        IF NOT stCmd.bEnable THEN
            // Route disable through STOPPING so MC_Stop runs first. If torque was
            // applied the axis is still in CST (torque) mode after Stop Torque;
            // MC_Stop performs the CST->position changeover and decelerates to a
            // real standstill BEFORE MC_Power drops. Withdrawing controller enable
            // straight from CST tripped NC 0x4260 (enable removed while the axis
            // was still positioning). STOPPING -> fbStop.Done -> DISABLED (SEL on
            // bEnable). Brief position hold during the decel, then power-off leaves
            // the motor free. (MOVING already disables via STOPPING; this makes
            // READY consistent. A normal idle disable just no-op-stops through it.)
            eState := E_MotorState.STOPPING;
        ELSIF fbPower.Error THEN
            eState := E_MotorState.ERROR;
        ELSIF rtStop.Q THEN
            eState := E_MotorState.STOPPING;
        ELSIF rtHome.Q THEN
            eState := E_MotorState.HOMING;
        ELSIF rtExecuteMove.Q THEN
            bMoveLatch := TRUE;
            eState     := E_MotorState.MOVING;
        END_IF

    E_MotorState.MOVING:
        IF NOT stCmd.bEnable OR rtStop.Q THEN
            bMoveLatch := FALSE;
            eState     := E_MotorState.STOPPING;

        ELSIF stCmd.eControlMode = E_ControlMode.POSITION THEN
            IF stCmd.bRelative THEN
                IF fbMoveRel.Busy  THEN bMoveLatch := FALSE; END_IF
                IF fbMoveRel.Done  THEN eState := E_MotorState.READY; END_IF
                IF fbMoveRel.Error THEN eState := E_MotorState.ERROR; END_IF
            ELSE
                IF fbMoveAbs.Busy  THEN bMoveLatch := FALSE; END_IF
                IF fbMoveAbs.Done  THEN eState := E_MotorState.READY; END_IF
                IF fbMoveAbs.Error THEN eState := E_MotorState.ERROR; END_IF
            END_IF

        ELSIF stCmd.eControlMode = E_ControlMode.VELOCITY THEN
            IF stCmd.fTargetVelocity <> fPrevVelocity THEN
                fPrevVelocity := stCmd.fTargetVelocity;
                bMoveLatch    := TRUE;
            END_IF
            IF fbMoveVel.Busy  THEN bMoveLatch := FALSE; END_IF
            IF fbMoveVel.Error THEN eState := E_MotorState.ERROR; END_IF

        ELSE
            eState := E_MotorState.READY;
        END_IF

    E_MotorState.STOPPING:
        IF fbStop.Error THEN
            eState := E_MotorState.ERROR;
        ELSIF fbStop.Done THEN
            eState := SEL(stCmd.bEnable, E_MotorState.DISABLED, E_MotorState.READY);
        END_IF

    E_MotorState.HOMING:
        fbHome(Axis := Axis, Execute := TRUE, HomingMode := MC_DefaultHoming);
        IF fbHome.Error THEN
            eState := E_MotorState.ERROR;
        ELSIF fbHome.Done THEN
            stStatus.bHomingDone := TRUE;
            eState               := E_MotorState.READY;
        END_IF

    E_MotorState.ERROR:
        IF rtResetError.Q THEN
            // Sequenced recovery: clear the DRIVE fault first (SoE S-0-0099),
            // give the drive a settle gap, THEN reset the NC axis against the
            // healthy drive. Sequenced on COMPLETION (Busy/Done), not timers.
            bSoeResetExec := TRUE;
            nResetStage   := 1;
            eState        := E_MotorState.RESETTING;
        END_IF

    E_MotorState.RESETTING:
        // Whole-sequence watchdog: if any stage hangs (e.g. a latch that never
        // clears), give up and go BACK TO ERROR — visible failure, another
        // reset press retries. Without this a stuck stage is unrecoverable
        // until a PLC restart.
        tonResetGuard(IN := TRUE, PT := T_RESET_GUARD);
        IF tonResetGuard.Q THEN
            tonResetGuard(IN := FALSE);
            bSoeResetExec := FALSE;
            bNcResetExec  := FALSE;
            nResetStage   := 0;
            eState        := E_MotorState.ERROR;
        END_IF
        CASE nResetStage OF
            1:  // SoE drive reset running — the latch self-clears when the
                // FB's Busy falls (done) or it errors/times out (10 s)
                IF NOT bSoeResetExec THEN
                    tonSettle(IN := FALSE);
                    nResetStage := 2;
                END_IF
            2:  // settle: let the drive's state machine come back up before
                // the NC touches it
                tonSettle(IN := TRUE, PT := T_RESET_SETTLE);
                IF tonSettle.Q THEN
                    tonSettle(IN := FALSE);
                    bNcResetExec := TRUE;
                    nResetStage  := 3;
                END_IF
            3:  // NC axis reset — latch self-clears on Done/Error
                IF NOT bNcResetExec THEN
                    tonResetGuard(IN := FALSE);
                    stStatus.bError   := FALSE;
                    stStatus.nErrorID := 0;
                    nResetStage       := 0;
                    eState            := E_MotorState.DISABLED;
                END_IF
        END_CASE

END_CASE

//----------------------------------------------------------------------
// STATUS OUTPUTS
//----------------------------------------------------------------------
stStatus.eState       := eState;
stStatus.eControlMode := stCmd.eControlMode;
stStatus.nResetStage  := nResetStage;
stStatus.bEnabled     := fbPower.Status;
stStatus.bMoving      := fbMoveAbs.Busy OR fbMoveRel.Busy OR fbMoveVel.Busy;
stStatus.bAtTarget    := fbMoveAbs.Done OR fbMoveRel.Done OR fbMoveVel.InVelocity;
// Error status sourced from the NC axis ErrorCode — the authoritative, PERSISTENT
// fault: set on any axis fault and HELD until MC_Reset. The MC-block .Error outputs
// are transient (they clear the moment a block's Execute drops or the axis
// disables), so the old MC-block-only bError usually went FALSE before the app
// polled and the error never reached the GUI (nErrorID lingered with bError=FALSE).
// Keep the block errors OR'd in; fall back to their ErrorID only when the axis has
// no code of its own; clear when truly error-free so a stale code can't linger.
stStatus.bError := (Axis.NcToPlc.ErrorCode <> 0)
                OR fbPower.Error   OR fbMoveAbs.Error OR fbMoveRel.Error
                OR fbMoveVel.Error OR fbStop.Error    OR fbHome.Error;

IF Axis.NcToPlc.ErrorCode <> 0 THEN
    stStatus.nErrorID := Axis.NcToPlc.ErrorCode;
ELSIF stStatus.bError THEN
    stStatus.nErrorID := SEL(fbPower.Error,   0, fbPower.ErrorID)
                       + SEL(fbMoveAbs.Error, 0, fbMoveAbs.ErrorID)
                       + SEL(fbMoveRel.Error, 0, fbMoveRel.ErrorID)
                       + SEL(fbMoveVel.Error, 0, fbMoveVel.ErrorID)
                       + SEL(fbStop.Error,    0, fbStop.ErrorID)
                       + SEL(fbHome.Error,    0, fbHome.ErrorID);
ELSE
    stStatus.nErrorID := 0;
END_IF

stStatus.fActPosition := Axis.NcToPlc.ActPos;
stStatus.fActVelocity := Axis.NcToPlc.ActVelo;
stStatus.fActTorque   := INT_TO_LREAL(nActTorque_Raw) / 10.0;
stStatus.nTimestamp   := ULINT_TO_UDINT(F_GetSystemTime() / 10000);

END_FUNCTION_BLOCK

// ---- POUs/FB_TorqueControl.TcPOU
FUNCTION_BLOCK FB_TorqueControl
VAR_IN_OUT
    Axis            : AXIS_REF;         // Must be VAR_IN_OUT — passed by reference
END_VAR

VAR_INPUT
    stCmd           : ST_MotorCommand;  // Read from GVL_Commands
    bAxisReady      : BOOL;             // gate: only stream torque while the axis is READY
END_VAR

VAR_OUTPUT
    stStatus        : ST_MotorStatus;   // Written to GVL_Status
END_VAR

VAR
    fbTorqueCtrl    : MC_TorqueControl;
    rtExecute       : R_TRIG;
END_VAR

// Rising edge on bTorqueExecute triggers MC_TorqueControl
rtExecute(CLK := stCmd.bTorqueExecute);

// Gate Execute on READY: torque must never be commanded on a DISABLED/ERROR/
// RESETTING axis. This also drops Execute on a fault (READY->ERROR), which
// clears MC_TorqueControl's latched Error, and prevents the reset "bounce"
// where torque errors on the just-disabled axis and re-stamps the fault.
fbTorqueCtrl(
    Axis              := Axis,
    Execute           := stCmd.bTorqueExecute AND bAxisReady,
    ContinuousUpdate  := TRUE,
    Relative          := FALSE,
    Torque            := stCmd.fTargetTorque,
    TorqueRamp        := stCmd.fTorqueRamp,
    VelocityLimitHigh := stCmd.fTorqueVelLimitHigh,
    VelocityLimitLow  := stCmd.fTorqueVelLimitLow,
    BufferMode        := MC_Aborting
);

// Write ONLY torque fields back — do not overwrite position/velocity status
stStatus.bTorqueActive   := fbTorqueCtrl.Active;
stStatus.bTorqueInTorque := fbTorqueCtrl.InTorque;

// Reflect the LIVE torque-FB error. This was set-only (no ELSE), so once a
// torque fault set bError it stayed latched forever and PRG_Motion's set-only
// copy re-stamped it onto the status mirror every scan — the motor recovered
// but bError/nErrorID never cleared. With Execute gated off on !READY, a reset
// clears MC_TorqueControl.Error and this ELSE then clears the mirror. A REAL,
// persistent torque fault keeps fbTorqueCtrl.Error TRUE, so it is not masked.
IF fbTorqueCtrl.Error THEN
    stStatus.bError   := TRUE;
    stStatus.nErrorID := fbTorqueCtrl.ErrorId;
ELSE
    stStatus.bError   := FALSE;
    stStatus.nErrorID := 0;
END_IF

END_FUNCTION_BLOCK

// ---- POUs/FB_IOHandler.TcPOU
FUNCTION_BLOCK FB_IOHandler
VAR_INPUT
    // Raw digital input byte — link this to your EL1008 terminal in XAE
    nRawDigitalIn   : BYTE;

    // Raw analog input values — link to EL3002 channels in XAE
    nRawAnalogIn_Ch1 : INT;
    nRawAnalogIn_Ch2 : INT;

    // Analog scaling — set once from MAIN or leave as defaults
    fAnalogIn_Scale_Ch1  : LREAL := 10.0;   // full-scale [V or mA]
    fAnalogIn_Scale_Ch2  : LREAL := 10.0;
    fAnalogOut_Scale_Ch1 : LREAL := 10.0;
    fAnalogOut_Scale_Ch2 : LREAL := 10.0;
END_VAR

VAR_OUTPUT
    // Packed digital output byte — link this to your EL2008 terminal in XAE
    nRawDigitalOut  : BYTE;

    // Raw analog output values — link to EL4002 channels in XAE
    nRawAnalogOut_Ch1 : INT;
    nRawAnalogOut_Ch2 : INT;
END_VAR

VAR_IN_OUT
    // Shared IO struct — same instance passed in from MAIN and GVL_IO
    stIO : ST_IOData;
END_VAR

//======================================================================
// DIGITAL INPUTS — unpack raw byte into named booleans
//======================================================================
stIO.bDI_EmergencyStop  := nRawDigitalIn.0;
stIO.bDI_HomeSensor_M1  := nRawDigitalIn.1;
stIO.bDI_HomeSensor_M2  := nRawDigitalIn.2;
stIO.bDI_LimitPos_M1    := nRawDigitalIn.3;
stIO.bDI_LimitNeg_M1    := nRawDigitalIn.4;
stIO.bDI_LimitPos_M2    := nRawDigitalIn.5;
stIO.bDI_LimitNeg_M2    := nRawDigitalIn.6;
stIO.bDI_UserInput1     := nRawDigitalIn.7;

// Mirror raw byte for Python diagnostics
stIO.nDigitalInputs     := nRawDigitalIn;

//======================================================================
// ANALOG INPUTS — scale INT [-32768..32767] → engineering units
// Formula: value = (raw / 32767.0) * full_scale
//======================================================================
stIO.fAnalogIn_Ch1      := (INT_TO_LREAL(nRawAnalogIn_Ch1) / 32767.0)
                            * fAnalogIn_Scale_Ch1;
stIO.fAnalogIn_Ch2      := (INT_TO_LREAL(nRawAnalogIn_Ch2) / 32767.0)
                            * fAnalogIn_Scale_Ch2;
stIO.nAnalogIn_Raw_Ch1  := nRawAnalogIn_Ch1;
stIO.nAnalogIn_Raw_Ch2  := nRawAnalogIn_Ch2;

//======================================================================
// DIGITAL OUTPUTS — pack named booleans into raw byte for EL2008
//======================================================================
nRawDigitalOut.0 := stIO.bDO_BrakeRelease_M1;
nRawDigitalOut.1 := stIO.bDO_BrakeRelease_M2;
nRawDigitalOut.2 := stIO.bDO_StatusLED_Green;
nRawDigitalOut.3 := stIO.bDO_StatusLED_Red;
nRawDigitalOut.4 := stIO.bDO_UserOutput1;
nRawDigitalOut.5 := stIO.bDO_UserOutput2;

// Mirror packed byte back into struct for Python readback
stIO.nDigitalOutputs    := nRawDigitalOut;

//======================================================================
// ANALOG OUTPUTS — scale engineering units → INT [-32767..32767]
// Formula: raw = CLAMP(value / full_scale, -1.0, 1.0) * 32767
// Python writes fAnalogOut_Ch1/2 into GVL_IO.stIO, FB reads them here
//======================================================================
stIO.nAnalogOut_Raw_Ch1 := LREAL_TO_INT(
    LIMIT(-32767.0,
          (stIO.fAnalogOut_Ch1 / fAnalogOut_Scale_Ch1) * 32767.0,
          32767.0));

stIO.nAnalogOut_Raw_Ch2 := LREAL_TO_INT(
    LIMIT(-32767.0,
          (stIO.fAnalogOut_Ch2 / fAnalogOut_Scale_Ch2) * 32767.0,
          32767.0));

nRawAnalogOut_Ch1 := stIO.nAnalogOut_Raw_Ch1;
nRawAnalogOut_Ch2 := stIO.nAnalogOut_Raw_Ch2;

END_FUNCTION_BLOCK

// ---- POUs/FB_EncoderHandler.TcPOU
FUNCTION_BLOCK FB_EncoderHandler
VAR_IN_OUT
    stEncoder           : ST_EncoderData;
END_VAR

VAR_INPUT
    fCountsPerUnit      : LREAL := 1.0;
END_VAR

VAR
    nStatusWord_Raw      AT %I* : WORD;
    nCounterValue_Raw    AT %I* : DWORD;
    nFrequencyValue_Raw  AT %I* : DWORD;
    nState_Raw           AT %I* : BYTE;

    nSetCounterValue_Raw AT %Q* : DWORD;
    nControlWord_Raw     AT %Q* : WORD;

    rtSetCounter        : R_TRIG;
    rtZeroPosition      : R_TRIG;
END_VAR

//----------------------------------------------------------------------
// READ INPUTS
//----------------------------------------------------------------------
stEncoder.nStatusWord     := nStatusWord_Raw;
stEncoder.nCounterValue   := nCounterValue_Raw;
stEncoder.nFrequencyValue := nFrequencyValue_Raw;
stEncoder.nState          := nState_Raw;

stEncoder.bInputA           := nStatusWord_Raw.0;
stEncoder.bInputB           := nStatusWord_Raw.1;
stEncoder.bInputC           := nStatusWord_Raw.2;
stEncoder.bCounterUnderflow := nStatusWord_Raw.4;
stEncoder.bCounterOverflow  := nStatusWord_Raw.5;
stEncoder.bLatchValid       := nStatusWord_Raw.8;
stEncoder.bError            := nStatusWord_Raw.14;

IF fCountsPerUnit <> 0 THEN
    stEncoder.fPosition := DWORD_TO_LREAL(nCounterValue_Raw) / fCountsPerUnit;
END_IF

//----------------------------------------------------------------------
// WRITE OUTPUTS
//----------------------------------------------------------------------
rtSetCounter  (CLK := stEncoder.bSetCounter);
rtZeroPosition(CLK := stEncoder.bZeroPosition);

IF rtZeroPosition.Q THEN
    stEncoder.nSetCounterValue := 0;
    nSetCounterValue_Raw       := 0;
    nControlWord_Raw.2         := TRUE;   // bit 2 = 0x7000:03 Set counter
ELSIF rtSetCounter.Q THEN
    nSetCounterValue_Raw       := stEncoder.nSetCounterValue;
    nControlWord_Raw.2         := TRUE;
ELSE
    nControlWord_Raw.2         := FALSE;
END_IF

END_FUNCTION_BLOCK

// ---- POUs/FB_AnalogInHandler.TcPOU
FUNCTION_BLOCK FB_AnalogInHandler
VAR_IN_OUT
    stAnalogIn      : ST_AnalogInData;  // Shared with GVL_AnalogIn
END_VAR

VAR
    //--- EL3702 PDO inputs — oversampling x5 per channel ---
    // Each sample is a signed INT [-32768 to 32767]
    // AT %I* — linked in XAE instance tree to EL3702 PDO channels
    nCh1_S1     AT %I* : INT;   // Ch1 sample 1
    nCh1_S2     AT %I* : INT;   // Ch1 sample 2
    nCh1_S3     AT %I* : INT;   // Ch1 sample 3
    nCh1_S4     AT %I* : INT;   // Ch1 sample 4
    nCh1_S5     AT %I* : INT;   // Ch1 sample 5

    nCh2_S1     AT %I* : INT;   // Ch2 sample 1
    nCh2_S2     AT %I* : INT;   // Ch2 sample 2
    nCh2_S3     AT %I* : INT;   // Ch2 sample 3
    nCh2_S4     AT %I* : INT;   // Ch2 sample 4
    nCh2_S5     AT %I* : INT;   // Ch2 sample 5

    //--- Internal ---
    fCh1_Sum    : LREAL;
    fCh2_Sum    : LREAL;
    fScale      : LREAL;
END_VAR

//----------------------------------------------------------------------
// STORE RAW SAMPLES INTO STRUCT
//----------------------------------------------------------------------
stAnalogIn.nCh1_Sample[1] := nCh1_S1;
stAnalogIn.nCh1_Sample[2] := nCh1_S2;
stAnalogIn.nCh1_Sample[3] := nCh1_S3;
stAnalogIn.nCh1_Sample[4] := nCh1_S4;
stAnalogIn.nCh1_Sample[5] := nCh1_S5;

stAnalogIn.nCh2_Sample[1] := nCh2_S1;
stAnalogIn.nCh2_Sample[2] := nCh2_S2;
stAnalogIn.nCh2_Sample[3] := nCh2_S3;
stAnalogIn.nCh2_Sample[4] := nCh2_S4;
stAnalogIn.nCh2_Sample[5] := nCh2_S5;

//----------------------------------------------------------------------
// OVERSAMPLING PROCESSING — average 5 samples per channel
// Scale: INT [-32768..32767] → voltage [-fFullScale..+fFullScale]
// Formula: V = (avg_raw / 32767.0) * fFullScale
//----------------------------------------------------------------------
fScale := stAnalogIn.fFullScale / 32767.0;

fCh1_Sum := INT_TO_LREAL(nCh1_S1)
           + INT_TO_LREAL(nCh1_S2)
           + INT_TO_LREAL(nCh1_S3)
           + INT_TO_LREAL(nCh1_S4)
           + INT_TO_LREAL(nCh1_S5);

fCh2_Sum := INT_TO_LREAL(nCh2_S1)
           + INT_TO_LREAL(nCh2_S2)
           + INT_TO_LREAL(nCh2_S3)
           + INT_TO_LREAL(nCh2_S4)
           + INT_TO_LREAL(nCh2_S5);

stAnalogIn.fCh1_Voltage := (fCh1_Sum / 5.0) * fScale;
stAnalogIn.fCh2_Voltage := (fCh2_Sum / 5.0) * fScale;

END_FUNCTION_BLOCK

// ---- POUs/FB_MenteeMotorHandler.TcPOU
FUNCTION_BLOCK FB_MenteeMotorHandler
VAR_IN_OUT
    stCmd               : ST_MenteeMotorCmd;    // From GVL_MenteeMotor
    stStatus            : ST_MenteeMotorStatus; // To GVL_MenteeMotor
END_VAR

VAR
    //--- RxPDO outputs — AT %Q* — link to device 0x7000 PDOs in XAE ---
    q_kp                    AT %Q* : REAL;  // 0x7000:01 kp
    q_kd                    AT %Q* : REAL;  // 0x7000:02 kd
    q_p_des                 AT %Q* : REAL;  // 0x7000:03 p_des
    q_v_des                 AT %Q* : REAL;  // 0x7000:04 v_des
    q_torque_feed_forward   AT %Q* : REAL;  // 0x7000:05 torque_feed_forward
    q_max_torque            AT %Q* : REAL;  // 0x7000:06 max_torque

    //--- TxPDO inputs — AT %I* — link to device 0x6000 PDOs in XAE ---
    i_general_error_bits    AT %I* : BYTE;  // 0x6000:01 general_error_bits
    i_categorial_error_bits AT %I* : BYTE;  // 0x6000:02 categorial_error_bits
    i_motor_temp            AT %I* : BYTE;  // 0x6000:03 motor_temp
    i_theta                 AT %I* : REAL;  // 0x6000:04 theta
    i_d_theta               AT %I* : REAL;  // 0x6000:05 d_theta
    i_measured_torque       AT %I* : REAL;  // 0x6000:06 measured_torque
    i_motor_torque_pi_in    AT %I* : REAL;  // 0x6000:07 motor_torque_pi_in
    i_p_des_echo            AT %I* : REAL;  // 0x6000:08 p_des_echo
END_VAR

//----------------------------------------------------------------------
// WRITE RxPDO — GVL_MenteeMotor.stCmd → device every cycle
//----------------------------------------------------------------------
q_kp                  := stCmd.kp;
q_kd                  := stCmd.kd;
q_p_des               := stCmd.p_des;
q_v_des               := stCmd.v_des;
q_torque_feed_forward := stCmd.torque_feed_forward;
q_max_torque          := stCmd.max_torque;

//----------------------------------------------------------------------
// READ TxPDO — device → GVL_MenteeMotor.stStatus every cycle
//----------------------------------------------------------------------
stStatus.general_error_bits    := i_general_error_bits;
stStatus.categorial_error_bits := i_categorial_error_bits;
stStatus.motor_temp            := i_motor_temp;
stStatus.theta                 := i_theta;
stStatus.d_theta               := i_d_theta;
stStatus.measured_torque       := i_measured_torque;
stStatus.motor_torque_pi_in    := i_motor_torque_pi_in;
stStatus.p_des_echo            := i_p_des_echo;

END_FUNCTION_BLOCK

// ---- POUs/FB_Slot2PipeHandler.TcPOU
// Generic slot-2 debug-PDO pipe (SLOT2_DEBUG_PDO_PROTOCOL.md) presented through the
// LEGACY contract: consumes/produces the same ST_MenteeMotorV32OsCmd / *OsStatus as the
// old fixed pipe, so everything above (profiles, CSV player, recorder, snapshot, app)
// keeps working unchanged. Three jobs:
//
//   1. BINDING ENGINE — on GVL_Slot2.bConfigure, walks ST_Slot2Cfg over the op/strobe
//      protocol: CLEAR_ALL, then BIND_MON_OUT per monitor lane and BIND_MON_IN per
//      inject slot (addr<>0 = used). One command per ~6 cycles; fault -> error + stop.
//   2. INJECT — while RUN, streams the 8 legacy command fields into inject slots 0..7
//      (values written by the slave to the bound RAM addrs every cycle):
//      0 impedance_p_des | 1 impedance_v_des | 2 impedance_kp | 3 impedance_kd |
//      4 impedance_torque_ff | 5 setpoint_position | 6 setpoint_velocity | 7 setpoint_current
//      (stCmd.nControlWord is IGNORED — FSM/mode go via FB_MenteeSdoCmd / SDO 0x2000.)
//   3. STATUS ADAPTER — fills ST_MenteeMotorV32OsStatus from the debug TxPDO:
//      discrete fsm/main/mode/errors (+ a SYNTHESIZED nStatusWord in the legacy bit
//      layout), and the aSamples[0..9] oversample view rebuilt from the monitor lanes
//      with sample_idx SYNTHESIZED from capture_count (0x0A, new FW semantics: value =
//      stamp of newest delivered sample) so the recorder's dedup/timing math is exact:
//        idx40(k) = (capture_count - (n-1-k)) * prescaler      [40 kHz-equivalent]
//
// >>> LINK IN XAE (new ESI, slot-2 0x1601/0x1A01): q_* -> 0x7001:01..10 entries,
//     i_* -> 0x6001:01..0B, i_samples -> 0x6001:0C..6F (multi-select -> array link). <<<
FUNCTION_BLOCK FB_Slot2PipeHandler
VAR_IN_OUT
    stCmd       : ST_MenteeMotorV32OsCmd;      // legacy command contract (setpoints used)
    stStatus    : ST_MenteeMotorV32OsStatus;   // legacy status contract (fully populated)
END_VAR
VAR
    stEmptySample   : ST_MenteeMotorV32OsSample;   // all-zero (never written)
    //--- RxPDO 0x1601 outputs — AT %Q* — link to box 0x7001 entries ---
    q_op        AT %Q* : UDINT;   // 0x7001:01
    q_slot      AT %Q* : UDINT;   // 0x7001:02
    q_size      AT %Q* : UDINT;   // 0x7001:03
    q_strobe    AT %Q* : UDINT;   // 0x7001:04
    q_prescaler AT %Q* : UDINT;   // 0x7001:05
    q_addr      AT %Q* : UDINT;   // 0x7001:06
    q_inject    AT %Q* : ARRAY[0..9] OF UDINT;   // 0x7001:07..10

    //--- TxPDO 0x1A01 inputs — AT %I* — link to box 0x6001 entries ---
    i_fsm_state       AT %I* : UDINT;   // 0x6001:01
    i_main_state      AT %I* : UDINT;   // 0x6001:02
    i_motion_mode     AT %I* : UDINT;   // 0x6001:03
    i_motor_enabled   AT %I* : UDINT;   // 0x6001:04
    i_general_error   AT %I* : UDINT;   // 0x6001:05
    i_categorial_error AT %I* : UDINT;  // 0x6001:06
    i_last_op         AT %I* : UDINT;   // 0x6001:07
    i_fault           AT %I* : UDINT;   // 0x6001:08
    i_sample_count    AT %I* : UDINT;   // 0x6001:09
    i_capture_count   AT %I* : UDINT;   // 0x6001:0A (capture counter, new FW semantics)
    i_var_count       AT %I* : UDINT;   // 0x6001:0B
    i_samples         AT %I* : ARRAY[0..99] OF UDINT;   // 0x6001:0C..6F (lane-major, [lane*10+k])

    //--- binding engine state ---
    rConfigure  : R_TRIG;
    rClearAll   : R_TRIG;
    eState      : BYTE;      // mirrors GVL_Slot2.nBindState: 0 idle|1 clear|2 bind|3 run|4 error
    nStep       : INT;       // walk: 0 CLEAR_ALL | 1..10 mon lanes 0..9 | 11..20 inj slots 0..9
    nPhase      : INT;       // per-command: 0 arm+strobe | 1 wait | 2 settle
    nWait       : INT;
    nOpSent     : UDINT;
    bClearOnly  : BOOL;            // bClearAll path: stop after CLEAR_ALL (don't bind)
    cfg         : ST_Slot2Cfg;     // latched on bConfigure (walk reads the latch)

    //--- adapters ---
    uW          : U_WordReal;
    nPre        : UDINT;     // effective prescaler (>=1)
    n           : UDINT;     // valid samples this cycle (0..10)
    k           : UDINT;
END_VAR
VAR CONSTANT
    BS_IDLE     : BYTE := 0;
    BS_CLEAR    : BYTE := 1;
    BS_BIND     : BYTE := 2;
    BS_RUN      : BYTE := 3;
    BS_ERROR    : BYTE := 4;
    OP_NOP      : UDINT := 0;
    OP_BIND_OUT : UDINT := 1;
    OP_BIND_IN  : UDINT := 2;
    OP_CLEAR_ALL: UDINT := 5;
    WAIT_CYCLES : INT := 5;    // cycles after strobe before checking fault (1 kHz bus, 4 kHz slave)
END_VAR

//----------------------------------------------------------------------
// CONFIGURE / CLEAR triggERS
//----------------------------------------------------------------------
rConfigure(CLK := GVL_Slot2.bConfigure);
rClearAll (CLK := GVL_Slot2.bClearAll);

IF rConfigure.Q THEN
    cfg    := GVL_Slot2.stCfg;      // latch — the walk must not see mid-write edits
    nStep  := 0;
    nPhase := 0;
    bClearOnly := FALSE;
    GVL_Slot2.bBindError  := FALSE;
    GVL_Slot2.nFailedSlot := 16#FF;
    // Reset the oversample view so no slot carries values bound to the PREVIOUS
    // lane selection (e.g. a dropped ELF debug var leaking into the new session).
    FOR k := 0 TO 9 DO
        stStatus.aSamples[k] := stEmptySample;
    END_FOR
    eState := BS_CLEAR;
ELSIF rClearAll.Q THEN
    nStep  := 0;
    nPhase := 0;
    bClearOnly := TRUE;             // CLEAR_ALL, then stop (idle)
    eState := BS_CLEAR;
END_IF

nPre := MAX(1, cfg.nPrescaler);
q_prescaler := nPre;

//----------------------------------------------------------------------
// BINDING ENGINE — one op/strobe command at a time
//----------------------------------------------------------------------
CASE eState OF

BS_CLEAR, BS_BIND:
    CASE nPhase OF
    0:  // arm the current command (strobe still low from the settle phase)
        IF eState = BS_CLEAR THEN
            q_op := OP_CLEAR_ALL; q_slot := 0; q_size := 0; q_addr := 0;
        ELSE
            // nStep 1..10 -> monitor lane (nStep-1); 11..20 -> inject slot (nStep-11)
            IF nStep <= 10 THEN
                q_op   := OP_BIND_OUT;
                q_slot := TO_UDINT(nStep - 1);
                q_size := cfg.aMonSize[nStep - 1];
                q_addr := cfg.aMonAddr[nStep - 1];
            ELSE
                q_op   := OP_BIND_IN;
                q_slot := TO_UDINT(nStep - 11);
                q_size := cfg.aInjSize[nStep - 11];
                q_addr := cfg.aInjAddr[nStep - 11];
            END_IF
        END_IF
        nOpSent  := q_op;
        q_strobe := 1;
        nWait    := 0;
        nPhase   := 1;

    1:  // rising edge fired — give the slave a few cycles, then check the echo
        nWait := nWait + 1;
        IF nWait >= WAIT_CYCLES THEN
            q_strobe := 0;
            IF (i_fault <> 0) OR (i_last_op <> nOpSent) THEN
                GVL_Slot2.bBindError  := TRUE;
                GVL_Slot2.nFailedSlot := TO_BYTE(nStep);
                eState := BS_ERROR;
            ELSE
                nPhase := 2;
                nWait  := 0;
            END_IF
        END_IF

    2:  // settle one cycle with strobe low, then advance to the next used entry
        nPhase := 0;
        REPEAT
            nStep := nStep + 1;
        UNTIL nStep > 20
           OR (nStep <= 10  AND cfg.aMonAddr[nStep - 1]  <> 0)
           OR (nStep >= 11 AND nStep <= 20 AND cfg.aInjAddr[nStep - 11] <> 0)
        END_REPEAT;
        IF eState = BS_CLEAR THEN
            // CLEAR done. bConfigure walk continues into BIND; bClearAll stops here.
            IF bClearOnly THEN
                eState := BS_IDLE;
            ELSIF nStep > 20 THEN
                eState := BS_RUN;       // nothing to bind (all addrs 0) — pipe runs bare
            ELSE
                eState := BS_BIND;
            END_IF
        ELSIF nStep > 20 THEN
            eState := BS_RUN;           // walk complete
        END_IF
    END_CASE

BS_RUN, BS_IDLE, BS_ERROR:
    q_op := OP_NOP; q_strobe := 0;

END_CASE

//----------------------------------------------------------------------
// INJECT — stream the legacy command fields into the bound write slots
//----------------------------------------------------------------------
IF eState = BS_RUN THEN
    // All 10 inject slots are written every cycle. Slots 2..7 are the default
    // command set (FW self-bound). Slots 0/1/8/9 are SPARE raw lanes: the app
    // streams bit-encoded values (via GVL_MenteeMotorV32_OS.stCmd.nRawInjectN)
    // for ELF-picked inject targets; copied VERBATIM (no float union) so integer
    // picks are not reinterpreted as floats. Unbound spares are ignored by the FW.
    q_inject[0] := stCmd.nRawInject0;                          // spare
    q_inject[1] := stCmd.nRawInject1;                          // spare
    uW.f := stCmd.impedance_kp;        q_inject[2] := uW.u;
    uW.f := stCmd.impedance_kd;        q_inject[3] := uW.u;
    uW.f := stCmd.impedance_torque_ff; q_inject[4] := uW.u;
    // Slots 5/6 fed MODE-AWARE (impedance_* in Impedance mode, else setpoint_*) —
    // the FW merged the twin pairs into one var each (target_p_des / v_des).
    IF i_motion_mode = 4 THEN          // Impedance mode -> the impedance_* fields
        uW.f := stCmd.impedance_p_des;   q_inject[5] := uW.u;   // -> target_p_des
        uW.f := stCmd.impedance_v_des;   q_inject[6] := uW.u;   // -> v_des
    ELSE                               // Position/Velocity/... -> the setpoint_* fields
        uW.f := stCmd.setpoint_position; q_inject[5] := uW.u;   // -> target_p_des
        uW.f := stCmd.setpoint_velocity; q_inject[6] := uW.u;   // -> v_des
    END_IF
    uW.f := stCmd.setpoint_current;    q_inject[7] := uW.u;
    q_inject[8] := stCmd.nRawInject8;                          // spare
    q_inject[9] := stCmd.nRawInject9;                          // spare
END_IF

//----------------------------------------------------------------------
// STATUS ADAPTER — legacy struct from the debug TxPDO
//----------------------------------------------------------------------
stStatus.nFsmState            := UDINT_TO_BYTE(i_fsm_state);
stStatus.nMainState           := UDINT_TO_BYTE(i_main_state);
stStatus.nOpMode              := UDINT_TO_BYTE(i_motion_mode);
stStatus.nGeneralErrorBits    := UDINT_TO_BYTE(i_general_error AND 16#FF);
stStatus.nCategorialErrorBits := UDINT_TO_BYTE(i_categorial_error AND 16#FF);
stStatus.bError               := (stStatus.nGeneralErrorBits <> 0)
                               OR (stStatus.nCategorialErrorBits <> 0);
// Synthesized legacy status word (MASTER_INTERFACE §4.4 layout) so recordings and any
// raw-word consumer decode exactly as before:
//   FSM[4:0] | main[8:5] | mode[11:9] | enabled[12] | (15:13 unused) | gen[23:16] | cat[31:24]
// Bits 15:13 used to carry the oversample GROUP_ID; that mechanism is gone (the
// ELF debug-var lanes replaced it), so they are simply left 0.
stStatus.nStatusWord :=
      (i_fsm_state AND 16#1F)
    + (i_main_state AND 16#0F)       * 16#20
    + (i_motion_mode AND 16#07)      * 16#200
    + (i_motor_enabled AND 16#01)    * 16#1000
    + (i_general_error AND 16#FF)    * 16#10000
    + (i_categorial_error AND 16#FF) * 16#1000000;

// Rolling counter: capture_count IS the new free-running counter (liveness = advancing).
stStatus.nSampleCount := i_capture_count;

// Oversample view: rebuild aSamples[] from the monitor lanes; sample_idx synthesized in
// 40 kHz units (stamp*prescaler) so the app/recorder timing math (idx/40kHz) is exact.
n := MIN(i_sample_count, 10);
IF eState = BS_RUN AND n > 0 THEN
    // Lanes 0/1/2 = theta/d_theta/iq -> w0/w1/w2 per sample;
    // lanes 3..9 = ELF-picked debug variables -> w3..w9. Every lane shares
    // the same capture index k (the FW samples all bound lanes on one
    // prescaler tick), so one aSamples[k] is one synchronized instant.
    FOR k := 0 TO n - 1 DO
        stStatus.aSamples[k].sample_idx := (i_capture_count - (n - 1 - k)) * nPre;
        stStatus.aSamples[k].w0 := i_samples[0*10 + k];
        stStatus.aSamples[k].w1 := i_samples[1*10 + k];
        stStatus.aSamples[k].w2 := i_samples[2*10 + k];
        stStatus.aSamples[k].w3 := i_samples[3*10 + k];
        stStatus.aSamples[k].w4 := i_samples[4*10 + k];
        stStatus.aSamples[k].w5 := i_samples[5*10 + k];
        stStatus.aSamples[k].w6 := i_samples[6*10 + k];
        stStatus.aSamples[k].w7 := i_samples[7*10 + k];
        stStatus.aSamples[k].w8 := i_samples[8*10 + k];
        stStatus.aSamples[k].w9 := i_samples[9*10 + k];
    END_FOR
    // Legacy invariant: slot 9 = the NEWEST sample (the app's live pos/vel/current
    // + liveness read aSamples[9]). Mirror the newest into EVERY unwritten slot
    // (n..9), not just slot 9: a slot that never refreshes would keep a stale
    // sample_idx from PLC start (raw 0) forever, and once the live index enters
    // the top quarter of u32 the recorder's wrap heuristic reads that stale 0 as
    // a 2^32 wrap EVERY frame — runaway timestamps + garbage rows. Mirrored
    // slots carry the newest stamp, so the recorder's monotonic-idx dedup drops
    // them exactly like the old slot-9 mirror.
    IF n < 10 THEN
        FOR k := n TO 9 DO
            stStatus.aSamples[k] := stStatus.aSamples[n - 1];
        END_FOR
    END_IF
    uW.u := i_samples[0*10 + (n-1)]; stStatus.fLatestPos     := uW.f;
    uW.u := i_samples[1*10 + (n-1)]; stStatus.fLatestVel     := uW.f;
    uW.u := i_samples[2*10 + (n-1)]; stStatus.fLatestCurrent := uW.f;
END_IF

//----------------------------------------------------------------------
// PIPE STATUS -> GVL (app diagnostics)
//----------------------------------------------------------------------
GVL_Slot2.nBindState    := eState;
GVL_Slot2.bPipeActive   := (eState = BS_RUN);
GVL_Slot2.nCaptureCount := i_capture_count;
GVL_Slot2.nVarCount     := i_var_count;
GVL_Slot2.nLastOp       := i_last_op;
GVL_Slot2.nFault        := i_fault;

END_FUNCTION_BLOCK

// ---- POUs/FB_MenteeSdoCmd.TcPOU
// CoE SDO command channel to the Mentee Motor Slave V3.2: writes one ec_command_id_e
// opcode byte to object 0x2000:01 (the slave's command interface — FSM/main/mode/
// enable; opcodes in cmd/cmd_handler.h). Replaces the legacy slot-2 control_word
// path: the generic debug RxPDO carries no control word.
//
// Driven via GVL_Slot2: app writes nSdoOpcode + pulses bSdoExecute; results come back
// on bSdoDone/bSdoError/nSdoErrId. One command in flight at a time.
//
// >>> LINK IN XAE: <Motor Slave box> > InfoData > AdsAddr  ->  stAdsAddr. <<<
// (EtherCAT master NetId + the slave's fixed address arrive automatically — no
// hardcoded NetId. Enable "Include ADS Address" in the slave's InfoData if hidden.)
FUNCTION_BLOCK FB_MenteeSdoCmd
VAR
    stAdsAddr    AT %I* : AMSADDR;      // Motor Slave InfoData.AdsAddr (NetId + port)

    fbSdoWrite   : FB_EcCoESdoWrite;
    rExec        : R_TRIG;
    byOpcode     : BYTE;                // latched opcode for the in-flight write
    bRunning     : BOOL;
    bPending     : BOOL;                // execute edge arrived while busy/cooling — run next
    bCooldown    : BOOL;                // one cycle with bExecute=FALSE so the FB re-arms
    sNetId       : T_AmsNetId;          // dotted string built from stAdsAddr.netId
    i            : INT;
END_VAR
VAR CONSTANT
    CMD_INDEX    : WORD := 16#2000;
    CMD_SUBINDEX : BYTE := 1;
END_VAR

// Build the master NetId string from the linked AMS address (e.g. '5.69.55.234.2.1').
// Manual concat -> no extra library dependency.
sNetId := '';
FOR i := 0 TO 5 DO
    sNetId := CONCAT(sNetId, BYTE_TO_STRING(stAdsAddr.netId[i]));
    IF i < 5 THEN
        sNetId := CONCAT(sNetId, '.');
    END_IF
END_FOR

rExec(CLK := GVL_Slot2.bSdoExecute);

// An execute edge while a write is in flight (or during the re-arm cycle) is
// LATCHED, not lost — it starts as soon as the FB has re-armed.
IF rExec.Q AND (bRunning OR bCooldown) THEN
    bPending := TRUE;
END_IF

// Start a new write on the rising edge (or a latched pending one) — only when idle
// AND after >=1 cycle with bExecute=FALSE (bCooldown) so the FB sees a clean edge.
IF (rExec.Q OR bPending) AND NOT bRunning AND NOT bCooldown THEN
    bPending          := FALSE;
    byOpcode          := GVL_Slot2.nSdoOpcode;
    GVL_Slot2.bSdoDone  := FALSE;
    GVL_Slot2.bSdoError := FALSE;
    GVL_Slot2.nSdoErrId := 0;
    bRunning          := TRUE;
END_IF

fbSdoWrite(
    sNetId     := sNetId,
    nSlaveAddr := stAdsAddr.port,       // slave's fixed EtherCAT address (from AdsAddr)
    nIndex     := CMD_INDEX,
    nSubIndex  := CMD_SUBINDEX,
    pSrcBuf    := ADR(byOpcode),
    cbBufLen   := 1,
    bExecute   := bRunning,
    tTimeout   := T#1S
);

// The FB raises bBusy on the same call that sees the bExecute rising edge, so once
// bRunning is set, "NOT bBusy" after the call above means the write finished.
bCooldown := FALSE;
IF bRunning AND NOT fbSdoWrite.bBusy THEN
    IF fbSdoWrite.bError THEN
        GVL_Slot2.bSdoError := TRUE;
        GVL_Slot2.nSdoErrId := fbSdoWrite.nErrId;
    ELSE
        GVL_Slot2.bSdoDone := TRUE;
    END_IF
    bRunning  := FALSE;                 // drop bExecute -> FB re-arms
    bCooldown := TRUE;                  // next cycle runs the FB with bExecute=FALSE first
END_IF

GVL_Slot2.bSdoBusy := bRunning OR bPending;

END_FUNCTION_BLOCK

// ---- POUs/FB_MenteeFoeFlash.TcPOU
// Flash a config.bin to the Mentee Motor Slave V3.2 over FoE, then persist it.
//
// Sequence (driven via GVL_MenteeFoe): on bExecute rising edge, with nLen>0 —
//   OPEN  -> FB_EcFoeOpen  (file "config.bin", write mode)
//   WRITE -> FB_EcFoeAccess (send aData[0..nLen-1] in one go)
//   CLOSE -> FB_EcFoeClose
//   SAVE  -> FB_EcCoESdoWrite 0x1010:01 = 0x65766173 ("save")  [auto, ONLY on a
//            validated download] -> firmware writes flash sector 7 + self-resets.
//
// The slave validates the 32-byte header + CRC32 during the FoE data phase; a bad
// file makes it return a FoE program-error, so a clean transfer (no bError AND
// cbDone == nLen) means received + validated + applied to RAM. The save is gated
// on that, so a failed download never commits to flash (bDownloadOk stays FALSE).
//
// >>> LINK IN XAE: <Motor Slave box> > InfoData > AdsAddr -> stAdsAddr. <<<
// Same AMS address as FB_MenteeSdoCmd (EtherCAT master NetId + slave fixed addr);
// FoE and CoE both use it. Enable "Include ADS Address" on the slave if hidden.
// Caller must ensure the motor is IDLE before pulsing bExecute (app enforces it).
FUNCTION_BLOCK FB_MenteeFoeFlash
VAR
    stAdsAddr AT %I* : AMSADDR;         // Motor Slave InfoData.AdsAddr (NetId + port)

    fbOpen       : FB_EcFoeOpen;
    fbAccess     : FB_EcFoeAccess;
    fbClose      : FB_EcFoeClose;
    fbSave       : FB_EcCoESdoWrite;
    rExec        : R_TRIG;
    sNetId       : T_AmsNetId;          // dotted string built from stAdsAddr.netId
    i            : INT;
    nSaveSig     : UDINT := 16#65766173;   // "save" (CoE Store Parameters signature)
    bPendErr     : BOOL;                // WRITE failed -> still CLOSE the port, then ERROR
    eState       : INT;
END_VAR
VAR CONSTANT
    ST_IDLE      : INT := 0;
    ST_OPEN      : INT := 1;
    ST_WRITE     : INT := 2;
    ST_CLOSE     : INT := 3;
    ST_SAVE      : INT := 4;
    ST_DONE      : INT := 5;
    ST_ERR       : INT := 6;
    CFG_FILE     : T_MaxString := 'config.bin';
    STORE_INDEX  : WORD := 16#1010;
    STORE_SUB    : BYTE := 1;
END_VAR

// Build the master NetId string from the linked AMS address (manual concat -> no
// extra library dependency), same as FB_MenteeSdoCmd.
sNetId := '';
FOR i := 0 TO 5 DO
    sNetId := CONCAT(sNetId, BYTE_TO_STRING(stAdsAddr.netId[i]));
    IF i < 5 THEN
        sNetId := CONCAT(sNetId, '.');
    END_IF
END_FOR

// Start on a rising edge, only when idle and there is data. Clear prior status.
rExec(CLK := GVL_MenteeFoe.bExecute);
IF rExec.Q AND (eState = ST_IDLE) AND (GVL_MenteeFoe.nLen > 0) THEN
    GVL_MenteeFoe.bDownloadOk := FALSE;
    GVL_MenteeFoe.bDone       := FALSE;
    GVL_MenteeFoe.bError      := FALSE;
    GVL_MenteeFoe.nErrId      := 0;
    GVL_MenteeFoe.nStage      := 0;
    bPendErr                  := FALSE;
    eState                    := ST_OPEN;
END_IF

// Call every sub-FB each cycle; bExecute is gated by the current state. Each
// Tc2_EtherCAT FB raises bBusy on the same call that sees the rising edge, so
// "state active AND NOT bBusy" reliably means that stage finished.
fbOpen(sNetId := sNetId, nPort := stAdsAddr.port, sPathName := CFG_FILE,
       dwPass := 0, eMode := eFoeMode_Write,
       bExecute := (eState = ST_OPEN), tTimeout := T#10S);

fbAccess(hFoe := fbOpen.hFoe, pBuffer := ADR(GVL_MenteeFoe.aData),
         cbBuffer := GVL_MenteeFoe.nLen,
         bExecute := (eState = ST_WRITE), tTimeout := T#20S);

fbClose(hFoe := fbOpen.hFoe, bExecute := (eState = ST_CLOSE), tTimeout := T#10S);

fbSave(sNetId := sNetId, nSlaveAddr := stAdsAddr.port,
       nIndex := STORE_INDEX, nSubIndex := STORE_SUB,
       pSrcBuf := ADR(nSaveSig), cbBufLen := 4,
       bExecute := (eState = ST_SAVE), tTimeout := T#5S);

CASE eState OF

ST_OPEN:
    IF NOT fbOpen.bBusy THEN
        IF fbOpen.bError THEN
            GVL_MenteeFoe.nStage := 1; GVL_MenteeFoe.nErrId := fbOpen.nErrId;
            eState := ST_ERR;                 // nothing opened -> no close needed
        ELSE
            eState := ST_WRITE;
        END_IF
    END_IF

ST_WRITE:
    IF NOT fbAccess.bBusy THEN
        IF fbAccess.bError OR (fbAccess.cbDone <> GVL_MenteeFoe.nLen) THEN
            bPendErr := TRUE;                 // still close the port, then report error
            GVL_MenteeFoe.nStage := 2;
            GVL_MenteeFoe.nErrId := fbAccess.nErrId;
        ELSE
            GVL_MenteeFoe.bDownloadOk := TRUE;   // received + validated by the slave
        END_IF
        eState := ST_CLOSE;
    END_IF

ST_CLOSE:
    IF NOT fbClose.bBusy THEN
        IF bPendErr THEN
            eState := ST_ERR;                 // the WRITE failed (nStage/nErrId set)
        ELSE
            // Download validated: the slave ACKed every byte (cbDone = nLen),
            // CRC-checked the payload and applied it to RAM. FoE has no protocol
            // file-end — the slave finalizes on the config.bin header size and ends
            // the session itself, so FB_EcFoeClose often returns a benign device
            // error (e.g. 0x700: no session to close). Close is best-effort cleanup;
            // proceed to save regardless of its result.
            eState := ST_SAVE;                // download OK -> auto-save
        END_IF
    END_IF

ST_SAVE:
    IF NOT fbSave.bBusy THEN
        IF fbSave.bError THEN
            GVL_MenteeFoe.nStage := 4; GVL_MenteeFoe.nErrId := fbSave.nErrId;
            eState := ST_ERR;
        ELSE
            GVL_MenteeFoe.bDone := TRUE;      // saved -> motor self-resets with the new config
            eState := ST_DONE;
        END_IF
    END_IF

ST_DONE:
    GVL_MenteeFoe.bError := FALSE;
    IF NOT GVL_MenteeFoe.bExecute THEN eState := ST_IDLE; END_IF   // re-arm on falling edge

ST_ERR:
    GVL_MenteeFoe.bError := TRUE;
    IF NOT GVL_MenteeFoe.bExecute THEN eState := ST_IDLE; END_IF

END_CASE

GVL_MenteeFoe.nState := eState;
GVL_MenteeFoe.bBusy  := (eState = ST_OPEN) OR (eState = ST_WRITE)
                        OR (eState = ST_CLOSE) OR (eState = ST_SAVE);

END_FUNCTION_BLOCK

// ---- POUs/FB_TrajectoryGen.TcPOU
// Generic 1 kHz motion-profile generator for the V3.2 motor. Evaluates the
// selected shape as value(t) online (no precomputed array) and streams it to
// the field PRG_Motion routes by nField. Shapes ported from the Cheetah
// ProfileGenerator: Sinusoidal / Trapezoidal / Step / S-Curve / Ramp, plus
// two point-to-point shapes (velocity-trapezoid displacement, planned by the
// app from v_max/a_max): P2P moves one leg and holds at the end; P2P_RT goes
// out and back (v = 0 at the turnaround), so repetitive reps chain without a
// jump. For both, fPeakValue is the SIGNED cruise velocity, fAccelTime/
// fSteadyTime/fDecelTime are the leg's segment times, and fStartValue is the
// ABSOLUTE anchor position the app planned from (exact landing on target).
//
// On Start the command is LATCHED into 'cfg' (a local copy of stTraj). The
// generator + the valueAt method read 'cfg' only -- so mid-run parameter
// changes are ignored, and the method never touches the VAR_IN_OUT (no C0371).
//
// Anchoring: for position-target fields (nField 0/1) the profile rides on the
// rotor's position captured at Start -> out = startPos + (value(t) - value(0)),
// so it begins exactly where the motor is (no jump). Velocity/current (2/3) use
// the value directly. Repetitive loops the whole profile (nReps; 0 = infinite),
// resting fRestS between reps.
FUNCTION_BLOCK FB_TrajectoryGen
VAR_IN_OUT
    stTraj          : ST_MenteeTrajCmd;
END_VAR
VAR_INPUT
    fMeasuredPos    : REAL;     // current measured output position [rad]
    fDt             : REAL;     // task cycle time [s]
    bStartSync      : BOOL;     // shared synchronized start (PRG_Motion gates with the Mentee enable)
    bStopSync       : BOOL;     // shared synchronized stop
END_VAR
VAR_OUTPUT
    bRunning        : BOOL;
    fSetpoint       : REAL;
    nFieldOut       : BYTE;     // LATCHED field of the running profile — route by
                                // this, not the live stTraj.nField, so an ADS
                                // reconfig mid-run can't misroute the output
END_VAR
VAR
    cfg             : ST_MenteeTrajCmd;   // latched command (read by body + valueAt)
    rStart          : R_TRIG;
    rStop           : R_TRIG;
    eState          : INT;      // see ST_* constants
    fElapsed        : REAL;     // time into the current run [s]
    fTotalDur       : REAL;     // total duration of one run [s]
    fStartPos       : REAL;     // anchor position (captured at Start)
    fValue0         : REAL;     // value(0) for anchoring
    bAnchor         : BOOL;     // position-target field -> anchor at current pos
    nRepDone        : UDINT;
    fRest           : REAL;     // rest countdown [s]
    fRaw            : REAL;
    bWasActive      : BOOL;
END_VAR
VAR CONSTANT
    ST_IDLE         : INT := 0;
    ST_RUN          : INT := 1;
    ST_REST         : INT := 2;
    ST_DONE         : INT := 3;
    SH_SINE         : BYTE := 0;
    SH_TRAP         : BYTE := 1;
    SH_STEP         : BYTE := 2;
    SH_SCURVE       : BYTE := 3;
    SH_RAMP         : BYTE := 4;
    SH_P2P          : BYTE := 5;
    SH_P2P_RT       : BYTE := 6;
END_VAR

rStart(CLK := stTraj.bStart OR bStartSync);
rStop(CLK := stTraj.bStop OR bStopSync);

// Stop -> hold current position (idle; PRG_Motion stops overriding the field).
IF rStop.Q THEN
    eState := ST_IDLE;
END_IF

// Start a new run -> latch the command into cfg; everything below reads cfg.
IF rStart.Q AND (stTraj.nShape <= SH_P2P_RT) AND (stTraj.nField <= 3) THEN
    cfg      := stTraj;
    nFieldOut := cfg.nField;
    fElapsed := 0.0;
    nRepDone := 0;
    // P2P ends AWAY from its start, so replaying it would jump the setpoint
    // back -> one-way moves are never repetitive (oscillation uses SH_P2P_RT).
    IF cfg.nShape = SH_P2P THEN
        cfg.bRepetitive := FALSE;
    END_IF
    // total duration of one run, per shape
    IF (cfg.nShape = SH_TRAP) OR (cfg.nShape = SH_SCURVE) OR (cfg.nShape = SH_P2P) THEN
        fTotalDur := cfg.fAccelTime + cfg.fSteadyTime + cfg.fDecelTime;
    ELSIF cfg.nShape = SH_P2P_RT THEN
        fTotalDur := 2.0 * (cfg.fAccelTime + cfg.fSteadyTime + cfg.fDecelTime);
    ELSE
        fTotalDur := cfg.fDuration;
    END_IF
    // position-target fields ride on the current position (no jump). The P2P
    // shapes anchor on the app's PLANNED start (fStartValue) instead, so the
    // move lands EXACTLY on the planned target; any drift accrued since
    // planning shows as a small initial step the servo absorbs (identical to
    // the app-side streamer these shapes replace).
    bAnchor := (cfg.nField = 0) OR (cfg.nField = 1);
    IF bAnchor THEN
        IF (cfg.nShape = SH_P2P) OR (cfg.nShape = SH_P2P_RT) THEN
            fStartPos := cfg.fStartValue;
        ELSE
            fStartPos := fMeasuredPos;
        END_IF
        fValue0   := valueAt(0.0);
    ELSE
        fStartPos := 0.0;
        fValue0   := 0.0;
    END_IF
    eState := ST_RUN;
END_IF

// "Active this cycle" is latched BEFORE transitions so the cycle that ends the
// run still writes the final value.
bWasActive := (eState = ST_RUN) OR (eState = ST_REST);

CASE eState OF

ST_RUN:
    fRaw := valueAt(fElapsed);
    IF bAnchor THEN
        stTraj.fSetpoint := fStartPos + (fRaw - fValue0);
    ELSE
        stTraj.fSetpoint := fRaw;
    END_IF
    fElapsed := fElapsed + fDt;
    IF fElapsed >= fTotalDur THEN
        // land on the exact end value
        fRaw := valueAt(fTotalDur);
        IF bAnchor THEN
            stTraj.fSetpoint := fStartPos + (fRaw - fValue0);
        ELSE
            stTraj.fSetpoint := fRaw;
        END_IF
        IF NOT cfg.bRepetitive THEN
            eState := ST_DONE;
        ELSE
            nRepDone := nRepDone + 1;
            IF (cfg.nReps > 0) AND (nRepDone >= cfg.nReps) THEN
                eState := ST_DONE;
            ELSE
                fRest  := cfg.fRestS;
                eState := ST_REST;
            END_IF
        END_IF
    END_IF

ST_REST:
    fRest := fRest - fDt;                   // hold last setpoint during the rest
    IF fRest <= 0.0 THEN
        fElapsed := 0.0;
        eState   := ST_RUN;
    END_IF

ST_DONE:
    ;                                       // hold fSetpoint

ST_IDLE:
    ;                                       // not running

END_CASE

stTraj.fElapsed := fElapsed;
bRunning        := bWasActive;
fSetpoint       := stTraj.fSetpoint;
stTraj.bRunning := bRunning;

// Signed displacement along one point-to-point velocity-trapezoid leg at
// time fT [s]: accelerate 0 -> fPeakValue over fAccelTime, cruise for
// fSteadyTime, decelerate back to 0 over fDecelTime. Clamps past the end, so
// leg(end) = fPeakValue * (fAccelTime/2 + fSteadyTime + fDecelTime/2) = the
// leg distance. Mirrors the app's TrapezoidProfile (trajectory.py) exactly.
METHOD p2pLeg : REAL
VAR_INPUT
    fT  : REAL;
END_VAR
VAR
    fTa : REAL;     // accel time [s]
    fTc : REAL;     // cruise time [s]
    fTd : REAL;     // decel time [s]
    fV  : REAL;     // signed cruise velocity
    fU  : REAL;
END_VAR
fTa := MAX(cfg.fAccelTime, 1E-6);
fTc := cfg.fSteadyTime;
fTd := MAX(cfg.fDecelTime, 1E-6);
fV  := cfg.fPeakValue;

IF fT <= 0.0 THEN
    p2pLeg := 0.0;
ELSIF fT < fTa THEN
    // accelerating: 1/2 * a * t^2 with a = fV / fTa
    p2pLeg := 0.5 * fV * fT * fT / fTa;
ELSIF fT < (fTa + fTc) THEN
    // cruising
    p2pLeg := fV * (0.5 * fTa + (fT - fTa));
ELSE
    // decelerating (clamped at the leg end)
    fU := fT - fTa - fTc;
    IF fU > fTd THEN fU := fTd; END_IF
    p2pLeg := fV * (0.5 * fTa + fTc + fU - 0.5 * fU * fU / fTd);
END_IF
END_METHOD

// Shape value at time fT [s] — closed-form, mirrors the Cheetah ProfileGenerator.
// Reads the latched 'cfg' (FB-local), never the VAR_IN_OUT.
METHOD valueAt : REAL
VAR_INPUT
    fT  : REAL;
END_VAR
VAR
    fU  : REAL;
END_VAR
VAR CONSTANT
    TWO_PI : REAL := 6.2831853;
END_VAR
CASE cfg.nShape OF

0:  // Sinusoidal: offset + A * sin(2*pi*f*t)
    valueAt := cfg.fOffset + cfg.fAmplitude * SIN(TWO_PI * cfg.fFrequency * fT);

1:  // Trapezoidal: ramp start->peak / hold / ramp peak->start
    IF fT < cfg.fAccelTime THEN
        valueAt := cfg.fStartValue
                 + (cfg.fPeakValue - cfg.fStartValue) * (fT / MAX(cfg.fAccelTime, 1E-6));
    ELSIF fT < (cfg.fAccelTime + cfg.fSteadyTime) THEN
        valueAt := cfg.fPeakValue;
    ELSE
        fU := (fT - cfg.fAccelTime - cfg.fSteadyTime) / MAX(cfg.fDecelTime, 1E-6);
        IF fU > 1.0 THEN fU := 1.0; END_IF
        valueAt := cfg.fPeakValue - (cfg.fPeakValue - cfg.fStartValue) * fU;
    END_IF

2:  // Step: start until step time, then end
    IF fT < cfg.fStepTime THEN
        valueAt := cfg.fStartValue;
    ELSE
        valueAt := cfg.fEndValue;
    END_IF

3:  // S-Curve: quintic smoothstep start->peak / hold / peak->start
    IF fT < cfg.fAccelTime THEN
        fU := fT / MAX(cfg.fAccelTime, 1E-6);
        valueAt := cfg.fStartValue
                 + (cfg.fPeakValue - cfg.fStartValue) * (fU*fU*fU*(10.0 + fU*(-15.0 + fU*6.0)));
    ELSIF fT < (cfg.fAccelTime + cfg.fSteadyTime) THEN
        valueAt := cfg.fPeakValue;
    ELSE
        fU := (fT - cfg.fAccelTime - cfg.fSteadyTime) / MAX(cfg.fDecelTime, 1E-6);
        IF fU > 1.0 THEN fU := 1.0; END_IF
        valueAt := cfg.fPeakValue
                 - (cfg.fPeakValue - cfg.fStartValue) * (fU*fU*fU*(10.0 + fU*(-15.0 + fU*6.0)));
    END_IF

4:  // Ramp: linear start->end over duration
    fU := fT / MAX(cfg.fDuration, 1E-6);
    IF fU > 1.0 THEN fU := 1.0; END_IF
    valueAt := cfg.fStartValue + (cfg.fEndValue - cfg.fStartValue) * fU;

5:  // P2P: one-way velocity-trapezoid displacement; ends at the leg distance
    valueAt := p2pLeg(fT);

6:  // P2P round trip: leg out, then the same leg mirrored back to the start
    fU := cfg.fAccelTime + cfg.fSteadyTime + cfg.fDecelTime;   // one leg [s]
    IF fT < fU THEN
        valueAt := p2pLeg(fT);
    ELSE
        valueAt := p2pLeg(fU) - p2pLeg(fT - fU);
    END_IF

ELSE
    valueAt := 0.0;
END_CASE
END_METHOD

END_FUNCTION_BLOCK

// ---- POUs/FB_LoadMotorProfile.TcPOU
// Load-motor (Beckhoff AX5000) motion-profile generator. Same online value(t)
// shapes as FB_TrajectoryGen, but applied in one of three DOMAINS (cfg.nDomain):
//
//   TORQUE   : fSetpoint is a torque % waveform. PRG_Motion streams it into
//              stMotorN_Cmd.fTargetTorque while bRunning; the existing
//              FB_TorqueControl (MC_TorqueControl, ContinuousUpdate) applies it.
//              No axis ownership change -> coexists with FB_MotorControl freely.
//
//   POSITION : fSetpoint is an absolute position [deg], anchored at the axis
//              actual position at Start (no jump). Fed via external setpoint
//              generation (MC_ExtSetPointGen*).
//
//   VELOCITY : fSetpoint is a velocity [deg/s] waveform, integrated to position
//              for the external-setpoint feed.
//
// IMPORTANT (POSITION/VELOCITY): this FB does NOT call MC_Power. The load motor
// must already be ENABLED (FB_MotorControl in READY) so FB_MotorControl stays the
// single power owner -> no MC_Power conflict. While the external generator is
// engaged FB_MotorControl's move FBs must stay idle (no MC_Move* executing); the
// app/sequencer guarantees this by not issuing moves during a profile.
//
// On Start the command is LATCHED into 'cfg'; valueAt + the body read cfg only.
FUNCTION_BLOCK FB_LoadMotorProfile
VAR_IN_OUT
    stProfile       : ST_LoadProfileCmd;
    Axis            : AXIS_REF;          // used for POSITION/VELOCITY external setpoint
END_VAR
VAR_INPUT
    fMeasuredPos    : LREAL;    // axis actual position [deg] (Axis.NcToPlc.ActPos, LREAL) for anchoring
    fDt             : REAL;     // task cycle time [s]
    bStartSync      : BOOL;     // shared synchronized start (self-gated by stProfile.bEnable)
    bStopSync       : BOOL;     // shared synchronized stop
END_VAR
VAR_OUTPUT
    bRunning        : BOOL;
    fSetpoint       : REAL;     // generated value, native units (% torque | deg | deg/s)
END_VAR
VAR
    cfg             : ST_LoadProfileCmd;  // latched command (read by body + valueAt)
    rStart          : R_TRIG;
    rStop           : R_TRIG;
    eState          : INT;
    fElapsed        : REAL;
    fTotalDur       : REAL;
    fStartPos       : LREAL;    // anchor (POSITION) / integrator base (VELOCITY) [deg] — LREAL to match the NC axis
    fValue0         : REAL;     // value(0) for POSITION anchoring (small shape value)
    bAnchor         : BOOL;     // POSITION domain -> anchor at current pos
    nRepDone        : UDINT;
    fRest           : REAL;
    fRaw            : REAL;
    bWasActive      : BOOL;
    fPosAccum       : LREAL;    // VELOCITY domain: integral of velocity [deg] — LREAL (large absolute)

    // external setpoint generation (POSITION / VELOCITY only)
    fbExtEnable     : MC_ExtSetPointGenEnable;
    fbExtDisable    : MC_ExtSetPointGenDisable;
    fbSyncPos       : MC_SetPosition;   // set := actual BEFORE engaging (see below)
    bSyncExec       : BOOL;     // latch: set-position sync requested / running
    bEnableExec     : BOOL;     // latch: ext-generator enable requested / running
    bWaitStill      : BOOL;     // latch: waiting for NC standstill before the sync
    tonStill        : TON;      // standstill-wait timeout (proceed anyway)
    rFeedOn         : R_TRIG;   // first feed cycle -> re-anchor at engagement
    bExtWant        : BOOL;     // this cycle wants the external generator engaged
    rExtOn          : R_TRIG;
    fExtOff         : F_TRIG;
    fExtPos         : LREAL;    // position fed to the generator [deg] — LREAL (NC interface)
    fExtVel         : LREAL;    // velocity fed [deg/s]
    fPrevExtPos     : LREAL;    // for POSITION numeric velocity feed-forward
    nExtDir         : DINT;     // 1 = +, -1 = -, 0 = standstill
END_VAR
VAR CONSTANT
    F_STILL_VELO    : LREAL := 1.0;    // NC standstill threshold [deg/s] before engaging
    T_STILL_TIMEOUT : TIME := T#2S;    // give up waiting for standstill -> proceed anyway
    ST_IDLE         : INT := 0;
    ST_RUN          : INT := 1;
    ST_REST         : INT := 2;
    ST_DONE         : INT := 3;
    DOM_TORQUE      : BYTE := 0;
    DOM_POSITION    : BYTE := 1;
    DOM_VELOCITY    : BYTE := 2;
    SH_SINE         : BYTE := 0;
    SH_TRAP         : BYTE := 1;
    SH_STEP         : BYTE := 2;
    SH_SCURVE       : BYTE := 3;
    SH_RAMP         : BYTE := 4;
END_VAR

// bStart (direct) OR a synchronized start gated by this profile's own bEnable.
rStart(CLK := stProfile.bStart OR (bStartSync AND stProfile.bEnable));
rStop (CLK := stProfile.bStop  OR bStopSync);

// Stop -> hold (idle; the external generator is disabled below on the falling edge).
IF rStop.Q THEN
    eState := ST_IDLE;
END_IF

// Start a new run -> latch the command into cfg; everything below reads cfg.
IF rStart.Q AND (stProfile.nShape <= SH_RAMP) AND (stProfile.nDomain <= DOM_VELOCITY) THEN
    cfg       := stProfile;
    fElapsed  := 0.0;
    nRepDone  := 0;
    fPosAccum := 0.0;
    // total duration of one run, per shape
    IF (cfg.nShape = SH_TRAP) OR (cfg.nShape = SH_SCURVE) THEN
        fTotalDur := cfg.fAccelTime + cfg.fSteadyTime + cfg.fDecelTime;
    ELSE
        fTotalDur := cfg.fDuration;
    END_IF
    // POSITION rides on the current axis position (no jump); VELOCITY integrates
    // from it; TORQUE is absolute.
    bAnchor := (cfg.nDomain = DOM_POSITION);
    IF (cfg.nDomain = DOM_POSITION) OR (cfg.nDomain = DOM_VELOCITY) THEN
        fStartPos := fMeasuredPos;
    ELSE
        fStartPos := 0.0;
    END_IF
    IF bAnchor THEN
        fValue0 := valueAt(0.0);
    ELSE
        fValue0 := 0.0;
    END_IF
    fPrevExtPos := fMeasuredPos;   // fresh velocity-FF seed (no spike from a prior run)
    eState := ST_RUN;
END_IF

// Latched BEFORE transitions so the cycle that ends the run still writes the value.
bWasActive := (eState = ST_RUN) OR (eState = ST_REST);

CASE eState OF

ST_RUN:
    // fSetpoint = the raw generated value (REAL telemetry / torque %). The absolute
    // POSITION/VELOCITY commands fed to the NC are built in LREAL below so a small
    // shape delta isn't swallowed when added to a large absolute axis position.
    fRaw := valueAt(fElapsed);
    stProfile.fSetpoint := fRaw;
    IF cfg.nDomain = DOM_VELOCITY THEN
        fPosAccum := fPosAccum + fRaw * fDt;
    END_IF
    fElapsed := fElapsed + fDt;
    IF fElapsed >= fTotalDur THEN
        // land on the exact end value
        fRaw := valueAt(fTotalDur);
        stProfile.fSetpoint := fRaw;
        IF NOT cfg.bRepetitive THEN
            eState := ST_DONE;
        ELSE
            nRepDone := nRepDone + 1;
            IF (cfg.nReps > 0) AND (nRepDone >= cfg.nReps) THEN
                eState := ST_DONE;
            ELSE
                fRest  := cfg.fRestS;
                eState := ST_REST;
            END_IF
        END_IF
    END_IF

ST_REST:
    fRest := fRest - fDt;                   // hold last value during the rest
    IF fRest <= 0.0 THEN
        fElapsed := 0.0;
        // VELOCITY rides on the position integral: re-anchor to the current actual
        // position and zero the accumulator each repeat, so any drift during the
        // rest is absorbed instead of compounding.
        IF cfg.nDomain = DOM_VELOCITY THEN
            fStartPos := fMeasuredPos;
            fPosAccum := 0.0;
        END_IF
        eState   := ST_RUN;
    END_IF

ST_DONE:
    ;                                       // hold fSetpoint

ST_IDLE:
    ;                                       // not running

END_CASE

//----------------------------------------------------------------------
// EXTERNAL SETPOINT GENERATION (POSITION / VELOCITY domains only).
// Engage on the first running cycle, feed each cycle while Enabled, disable when
// the run ends. TORQUE domain never touches the axis (PRG_Motion routes its value
// into stMotorN_Cmd.fTargetTorque).
//----------------------------------------------------------------------
bExtWant := ((cfg.nDomain = DOM_POSITION) OR (cfg.nDomain = DOM_VELOCITY))
            AND ((eState = ST_RUN) OR (eState = ST_REST));
rExtOn(CLK := bExtWant);
fExtOff(CLK := bExtWant);

// Engagement chain (POSITION/VELOCITY): scrub mailbox -> wait-standstill ->
// sync -> enable -> re-anchor at first feed.
// ROOT CAUSE of the F324 on profile sequences (bench-proven 2026-07-14):
// MC_ExtSetPointGenFeed writes a PERSISTENT PlcToNc image (ExtSetPos/Velo/
// Direction). Nothing cleared it after a run, so it kept the LAST run's
// sample armed (Direction<>0). At the next MC_ExtSetPointGenEnable the NC
// consumes that image in the 1..2-cycle window before the PLC can see
// Enabled and feed fresh values -> the drive command steps by the whole
// shaft displacement of the intervening torque run in ONE cycle -> F324
// (window ~5 deg / 250us on Axis 2). The scrub below (feed actual pos,
// vel 0, Direction 0 = "do not apply" while engagement is pending, plus a
// disarm sample at run end) closes that window. Standstill wait + sync stay
// as defense in depth against a stale NC setpoint.
IF rExtOn.Q THEN
    bWaitStill  := TRUE;                // stage 0: let residual creep die out
    bSyncExec   := FALSE;
    bEnableExec := FALSE;
    tonStill(IN := FALSE);
END_IF
IF fExtOff.Q THEN                       // run ended/stopped mid-sequence
    bWaitStill  := FALSE;
    bSyncExec   := FALSE;
    bEnableExec := FALSE;
    tonStill(IN := FALSE);
    // disarm the mailbox: leave the last commanded position with vel 0 and
    // Direction 0, so a later engagement can never replay this run's sample
    MC_ExtSetPointGenFeed(Position := fPrevExtPos, Velocity := 0.0,
                          Acceleration := 0.0, Direction := 0, Axis := Axis);
END_IF
// stage 0: NC-side standstill (position hold kills coast quickly); a
// SUSTAINED external drive can prevent it -> timeout proceeds anyway (the
// re-anchor below keeps the command step-free even then).
IF bWaitStill THEN
    tonStill(IN := TRUE, PT := T_STILL_TIMEOUT);
    IF (ABS(Axis.NcToPlc.ActVelo) <= F_STILL_VELO) OR tonStill.Q THEN
        tonStill(IN := FALSE);
        bWaitStill := FALSE;
        bSyncExec  := TRUE;             // stage 1: set := actual
    END_IF
END_IF
// stage 1: MC_SetPosition(set := actual) — moves a number, not the motor;
// no-op when set and actual already match.
fbSyncPos(Axis := Axis, Execute := bSyncExec,
          Position := fMeasuredPos, Mode := FALSE);
IF bSyncExec AND (fbSyncPos.Done OR fbSyncPos.Error) THEN
    bSyncExec := FALSE;
    IF bExtWant THEN
        bEnableExec := TRUE;            // stage 2: engage the generator
    END_IF
END_IF

fbExtEnable(
    Axis         := Axis,
    Execute      := bEnableExec,
    Position     := fMeasuredPos,
    PositionType := POSITIONTYPE_ABSOLUTE);
IF bEnableExec AND (fbExtEnable.Enabled OR fbExtEnable.Error) THEN
    bEnableExec := FALSE;               // one-shot: drop Execute once engaged
END_IF

// stage 3: re-anchor at the ACTUAL engagement instant. The start-edge anchor
// is stale by the standstill-wait + sync + enable cycles; on a shaft that
// crept meanwhile, feeding from the old anchor would step the command by the
// drift in one cycle (F324). Anchoring here makes the first command exactly
// the current position — step-free even on a still-moving shaft.
rFeedOn(CLK := fbExtEnable.Enabled AND bExtWant);
IF rFeedOn.Q THEN
    fStartPos   := fMeasuredPos;
    fValue0     := fRaw;        // shape continues from its current value
    fPosAccum   := 0.0;         // VELOCITY: restart the integral here
    fPrevExtPos := fMeasuredPos;
END_IF

IF fbExtEnable.Enabled AND bExtWant THEN
    IF cfg.nDomain = DOM_POSITION THEN
        // LREAL anchor + small REAL shape delta -> the delta survives the add
        fExtPos := fStartPos + (fRaw - fValue0);
        fExtVel := (fExtPos - fPrevExtPos) / MAX(fDt, 1E-6);   // numeric feed-forward
    ELSE
        // VELOCITY: position = start + integral; velocity = the value (0 in REST)
        fExtPos := fStartPos + fPosAccum;
        IF eState = ST_RUN THEN
            fExtVel := fRaw;
        ELSE
            fExtVel := 0.0;
        END_IF
    END_IF
    fPrevExtPos := fExtPos;

    IF   fExtVel > 0.0 THEN nExtDir := 1;
    ELSIF fExtVel < 0.0 THEN nExtDir := -1;
    ELSE                    nExtDir := 0;
    END_IF

    // Function: copies into the cyclic axis interface (fExtSetPos/Velo/Acc/Dir).
    MC_ExtSetPointGenFeed(
        Position     := fExtPos,
        Velocity     := fExtVel,
        Acceleration := 0.0,
        Direction    := nExtDir,
        Axis         := Axis);
ELSIF bExtWant THEN
    // engagement pending (standstill wait / sync / enable in flight): scrub
    // the mailbox every cycle so the NC's activation window can only ever
    // see (current actual position, vel 0, Direction 0 = do not apply)
    MC_ExtSetPointGenFeed(Position := fMeasuredPos, Velocity := 0.0,
                          Acceleration := 0.0, Direction := 0, Axis := Axis);
    fPrevExtPos := fMeasuredPos;
ELSE
    fPrevExtPos := fMeasuredPos;        // keep the derivative seed fresh while idle
END_IF

fbExtDisable(Axis := Axis, Execute := fExtOff.Q);

//----------------------------------------------------------------------
// STATUS
//----------------------------------------------------------------------
stProfile.fElapsed   := fElapsed;
bRunning             := bWasActive;
fSetpoint            := stProfile.fSetpoint;
stProfile.bRunning   := bRunning;
stProfile.bExtActive := fbExtEnable.Enabled;

// Shape value at time fT [s] — closed-form, mirrors FB_TrajectoryGen.valueAt.
// Reads the latched 'cfg' (FB-local), never the VAR_IN_OUT.
METHOD valueAt : REAL
VAR_INPUT
    fT  : REAL;
END_VAR
VAR
    fU  : REAL;
END_VAR
VAR CONSTANT
    TWO_PI : REAL := 6.2831853;
END_VAR
CASE cfg.nShape OF

0:  // Sinusoidal: offset + A * sin(2*pi*f*t)
    valueAt := cfg.fOffset + cfg.fAmplitude * SIN(TWO_PI * cfg.fFrequency * fT);

1:  // Trapezoidal: ramp start->peak / hold / ramp peak->start
    IF fT < cfg.fAccelTime THEN
        valueAt := cfg.fStartValue
                 + (cfg.fPeakValue - cfg.fStartValue) * (fT / MAX(cfg.fAccelTime, 1E-6));
    ELSIF fT < (cfg.fAccelTime + cfg.fSteadyTime) THEN
        valueAt := cfg.fPeakValue;
    ELSE
        fU := (fT - cfg.fAccelTime - cfg.fSteadyTime) / MAX(cfg.fDecelTime, 1E-6);
        IF fU > 1.0 THEN fU := 1.0; END_IF
        valueAt := cfg.fPeakValue - (cfg.fPeakValue - cfg.fStartValue) * fU;
    END_IF

2:  // Step: start until step time, then end
    IF fT < cfg.fStepTime THEN
        valueAt := cfg.fStartValue;
    ELSE
        valueAt := cfg.fEndValue;
    END_IF

3:  // S-Curve: quintic smoothstep start->peak / hold / peak->start
    IF fT < cfg.fAccelTime THEN
        fU := fT / MAX(cfg.fAccelTime, 1E-6);
        valueAt := cfg.fStartValue
                 + (cfg.fPeakValue - cfg.fStartValue) * (fU*fU*fU*(10.0 + fU*(-15.0 + fU*6.0)));
    ELSIF fT < (cfg.fAccelTime + cfg.fSteadyTime) THEN
        valueAt := cfg.fPeakValue;
    ELSE
        fU := (fT - cfg.fAccelTime - cfg.fSteadyTime) / MAX(cfg.fDecelTime, 1E-6);
        IF fU > 1.0 THEN fU := 1.0; END_IF
        valueAt := cfg.fPeakValue
                 - (cfg.fPeakValue - cfg.fStartValue) * (fU*fU*fU*(10.0 + fU*(-15.0 + fU*6.0)));
    END_IF

4:  // Ramp: linear start->end over duration
    fU := fT / MAX(cfg.fDuration, 1E-6);
    IF fU > 1.0 THEN fU := 1.0; END_IF
    valueAt := cfg.fStartValue + (cfg.fEndValue - cfg.fStartValue) * fU;

ELSE
    valueAt := 0.0;
END_CASE
END_METHOD

END_FUNCTION_BLOCK

// ---- POUs/FB_CsvPlayer.TcPOU
// Replays a CSV trajectory buffer (GVL_CsvProfile.stCsv) at the task rate. Each
// cycle it advances elapsed time, linearly interpolates BOTH channels at the same
// time index, and applies them -> the Mentee and the selected Beckhoff load motor
// stay synchronized (one player, one clock). Values are ABSOLUTE (no anchoring).
//
//   Mentee:   emits fMenteeOut; PRG_Motion routes it into the selected stCmd field
//             (setpoint_position | impedance_p_des | setpoint_velocity | setpoint_current).
//   Beckhoff: TORQUE   -> emits fLoadOut; PRG_Motion writes it to the selected
//                         motor's fTargetTorque (FB_TorqueControl streams it; the app
//                         must already be in torque mode).
//             POS/VEL  -> feeds the selected NC axis via external setpoint generation
//                         (MC_ExtSetPointGen*); the motor must be ENABLED/READY and not
//                         executing a move. VELOCITY integrates to position from the
//                         axis position captured at start.
//
// The scalar config is latched on the bStart edge; the sample arrays are read live
// (the app uploads them fully before pulsing bStart, and doesn't change them mid-run).
FUNCTION_BLOCK FB_CsvPlayer
VAR_IN_OUT
    stCsv           : ST_CsvProfile;
    AxisLoad1       : AXIS_REF;
    AxisLoad2       : AXIS_REF;
END_VAR
VAR_INPUT
    fLoad1Pos       : LREAL;    // Axis1.NcToPlc.ActPos [deg]
    fLoad2Pos       : LREAL;    // Axis2.NcToPlc.ActPos [deg]
    fDt             : REAL;     // task cycle time [s]
END_VAR
VAR_OUTPUT
    bRunning        : BOOL;
    fMenteeOut      : REAL;     // routed by PRG into the mentee field (while bRunning + enabled)
    fLoadOut        : REAL;     // routed by PRG into fTargetTorque (TORQUE domain, while bRunning + enabled)
END_VAR
VAR
    rStart          : R_TRIG;
    rStop           : R_TRIG;
    eState          : INT;
    fElapsed        : REAL;     // time into the current pass [s]
    fIdxR           : LREAL;    // fractional sample index
    iIdx            : DINT;
    fFrac           : REAL;
    fMenteeRaw      : REAL;
    fLoadRaw        : REAL;
    bWasActive      : BOOL;
    nRepDone        : UDINT;
    fRest           : REAL;

    // latched scalar config (read by the body; arrays read live from stCsv)
    nCountL         : UDINT;
    nLastIdx        : DINT;     // nCount-1
    fSampleDtL      : REAL;
    bMenteeEnL      : BOOL;
    nMenteeFieldL   : BYTE;
    bLoadEnL        : BOOL;
    nLoadMotorL     : BYTE;
    nLoadDomainL    : BYTE;
    bRepetitiveL    : BOOL;
    nRepsL          : UDINT;
    fRestSL         : REAL;

    // external setpoint generation (POSITION / VELOCITY) — instances per axis,
    // only the selected one is ever Execute'd.
    fbExt1On        : MC_ExtSetPointGenEnable;
    fbExt2On        : MC_ExtSetPointGenEnable;
    fbExt1Off       : MC_ExtSetPointGenDisable;
    fbExt2Off       : MC_ExtSetPointGenDisable;
    fbSync1         : MC_SetPosition;   // set := actual before engaging (F324/F321 guard)
    fbSync2         : MC_SetPosition;
    bSyncExec       : BOOL;     // latch: set-position sync requested / running
    bEnableExec     : BOOL;     // latch: ext-generator enable requested / running
    bSyncDone       : BOOL;
    bWaitStill      : BOOL;     // latch: waiting for NC standstill before the sync
    tonStill        : TON;      // standstill-wait timeout (proceed anyway)
    rFeedOn         : R_TRIG;   // first feed cycle -> re-anchor at engagement
    fActVelSel      : LREAL;    // selected load axis NC velocity [deg/s]
    rExtOn          : R_TRIG;
    fExtOff         : F_TRIG;
    bExtWant        : BOOL;
    bExtEnabled     : BOOL;
    fLoadStartPos   : LREAL;    // axis pos captured at start (VELOCITY integral base)
    fLoadPosAccum   : LREAL;    // VELOCITY: integral of velocity [deg]
    fExtPos         : LREAL;
    fExtVel         : LREAL;
    fPrevExtPos     : LREAL;
    nExtDir         : DINT;
END_VAR
VAR CONSTANT
    F_STILL_VELO    : LREAL := 1.0;    // NC standstill threshold [deg/s] before engaging
    T_STILL_TIMEOUT : TIME := T#2S;    // give up waiting for standstill -> proceed anyway
    ST_IDLE         : INT := 0;
    ST_RUN          : INT := 1;
    ST_REST         : INT := 2;
    ST_DONE         : INT := 3;
    DOM_TORQUE      : BYTE := 0;
    DOM_POSITION    : BYTE := 1;
    DOM_VELOCITY    : BYTE := 2;
END_VAR

rStart(CLK := stCsv.bStart);
rStop (CLK := stCsv.bStop);

IF rStop.Q THEN
    eState := ST_IDLE;
END_IF

// Start -> latch the scalar config; arrays are read live from stCsv.
IF rStart.Q AND (stCsv.nCount > 0) AND (stCsv.fSampleDt > 0.0) THEN
    nCountL       := stCsv.nCount;
    nLastIdx      := UDINT_TO_DINT(stCsv.nCount) - 1;
    fSampleDtL    := stCsv.fSampleDt;
    bMenteeEnL    := stCsv.bMenteeEnable;
    nMenteeFieldL := stCsv.nMenteeField;
    bLoadEnL      := stCsv.bLoadEnable;
    nLoadMotorL   := stCsv.nLoadMotor;
    nLoadDomainL  := stCsv.nLoadDomain;
    bRepetitiveL  := stCsv.bRepetitive;
    nRepsL        := stCsv.nReps;
    fRestSL       := stCsv.fRestS;
    fElapsed      := 0.0;
    nRepDone      := 0;
    fLoadPosAccum := 0.0;
    IF nLoadMotorL = 1 THEN fLoadStartPos := fLoad1Pos; ELSE fLoadStartPos := fLoad2Pos; END_IF
    fPrevExtPos   := fLoadStartPos;
    eState        := ST_RUN;
END_IF

bWasActive := (eState = ST_RUN) OR (eState = ST_REST);

CASE eState OF

ST_RUN:
    fIdxR := fElapsed / fSampleDtL;
    iIdx  := LREAL_TO_DINT(fIdxR);          // floor (fElapsed >= 0)
    IF iIdx >= nLastIdx THEN
        // reached the end of the table -> hold the last sample, then rep / done
        fMenteeRaw := stCsv.aMentee[nLastIdx];
        fLoadRaw   := stCsv.aLoad[nLastIdx];
        IF nLoadDomainL = DOM_VELOCITY THEN
            fLoadPosAccum := fLoadPosAccum + fLoadRaw * fDt;   // include the final sample
        END_IF
        IF NOT bRepetitiveL THEN
            eState := ST_DONE;
        ELSE
            nRepDone := nRepDone + 1;
            IF (nRepsL > 0) AND (nRepDone >= nRepsL) THEN
                eState := ST_DONE;
            ELSE
                fRest  := fRestSL;
                eState := ST_REST;
            END_IF
        END_IF
    ELSE
        fFrac      := LREAL_TO_REAL(fIdxR - DINT_TO_LREAL(iIdx));
        fMenteeRaw := stCsv.aMentee[iIdx] + fFrac * (stCsv.aMentee[iIdx + 1] - stCsv.aMentee[iIdx]);
        fLoadRaw   := stCsv.aLoad[iIdx]   + fFrac * (stCsv.aLoad[iIdx + 1]   - stCsv.aLoad[iIdx]);
        IF nLoadDomainL = DOM_VELOCITY THEN
            fLoadPosAccum := fLoadPosAccum + fLoadRaw * fDt;     // integrate velocity -> position
        END_IF
        fElapsed := fElapsed + fDt;
    END_IF

ST_REST:
    fRest := fRest - fDt;                   // hold last sample during the rest
    IF fRest <= 0.0 THEN
        fElapsed := 0.0;
        IF nLoadDomainL = DOM_VELOCITY THEN     // re-anchor so rest-drift doesn't compound
            fLoadStartPos := SEL(nLoadMotorL = 1, fLoad2Pos, fLoad1Pos);
            fLoadPosAccum := 0.0;
        END_IF
        eState := ST_RUN;
    END_IF

ST_DONE:
    ;                                       // hold last values

ST_IDLE:
    ;                                       // not running

END_CASE

//----------------------------------------------------------------------
// BECKHOFF external setpoint generation (POSITION / VELOCITY domains only).
//----------------------------------------------------------------------
bExtWant := bLoadEnL
            AND ((nLoadDomainL = DOM_POSITION) OR (nLoadDomainL = DOM_VELOCITY))
            AND ((eState = ST_RUN) OR (eState = ST_REST));
rExtOn(CLK := bExtWant);
fExtOff(CLK := bExtWant);

// Engagement chain: scrub mailbox -> wait-standstill -> sync -> enable ->
// re-anchor. See FB_LoadMotorProfile for the full F324 root-cause note:
// the PlcToNc ExtSetPos/Velo/Direction image persists between runs and the
// NC consumes it at generator activation before the first PLC feed; the
// Direction-0 scrub while engagement is pending closes that window.
IF rExtOn.Q THEN
    bWaitStill  := TRUE;                // stage 0: let the shaft settle first
    bSyncExec   := FALSE;
    bEnableExec := FALSE;
    tonStill(IN := FALSE);
END_IF
IF fExtOff.Q THEN                       // run ended/stopped mid-sequence
    bWaitStill  := FALSE;
    bSyncExec   := FALSE;
    bEnableExec := FALSE;
    tonStill(IN := FALSE);
    // disarm the mailbox: leave the last commanded position with vel 0 and
    // Direction 0, so a later engagement can never replay this run's sample
    IF nLoadMotorL = 1 THEN
        MC_ExtSetPointGenFeed(Position := fPrevExtPos, Velocity := 0.0,
                              Acceleration := 0.0, Direction := 0, Axis := AxisLoad1);
    ELSE
        MC_ExtSetPointGenFeed(Position := fPrevExtPos, Velocity := 0.0,
                              Acceleration := 0.0, Direction := 0, Axis := AxisLoad2);
    END_IF
END_IF

// stage 0: wait for NC standstill. After a high-amplitude TORQUE run the shaft
// is still creeping when the next profile starts; syncing/engaging on a moving
// shaft leaves the anchor stale by the time the first feed lands (F324).
// Timeout proceeds anyway so a slowly-drifting axis can't block the run.
IF bWaitStill THEN
    fActVelSel := SEL(nLoadMotorL = 1, AxisLoad2.NcToPlc.ActVelo, AxisLoad1.NcToPlc.ActVelo);
    tonStill(IN := TRUE, PT := T_STILL_TIMEOUT);
    IF (ABS(fActVelSel) <= F_STILL_VELO) OR tonStill.Q THEN
        tonStill(IN := FALSE);
        bWaitStill := FALSE;
        bSyncExec  := TRUE;
    END_IF
END_IF
fbSync1(Axis := AxisLoad1, Execute := bSyncExec AND (nLoadMotorL = 1),
        Position := fLoad1Pos, Mode := FALSE);
fbSync2(Axis := AxisLoad2, Execute := bSyncExec AND (nLoadMotorL = 2),
        Position := fLoad2Pos, Mode := FALSE);
bSyncDone := SEL(nLoadMotorL = 1,
                 fbSync2.Done OR fbSync2.Error,
                 fbSync1.Done OR fbSync1.Error);
IF bSyncExec AND bSyncDone THEN
    bSyncExec := FALSE;
    IF bExtWant THEN
        bEnableExec := TRUE;            // sync done -> now engage the generator
    END_IF
END_IF

fbExt1On(Axis := AxisLoad1, Execute := bEnableExec AND (nLoadMotorL = 1),
         Position := fLoad1Pos, PositionType := POSITIONTYPE_ABSOLUTE);
fbExt2On(Axis := AxisLoad2, Execute := bEnableExec AND (nLoadMotorL = 2),
         Position := fLoad2Pos, PositionType := POSITIONTYPE_ABSOLUTE);
bExtEnabled := SEL(nLoadMotorL = 1, fbExt2On.Enabled, fbExt1On.Enabled);  // selected axis
IF bEnableExec AND bExtEnabled THEN
    bEnableExec := FALSE;               // one-shot: drop Execute once engaged
END_IF

// stage 3: re-anchor at the ACTUAL engagement instant. The start-edge anchor
// is stale by the standstill-wait + sync + enable cycles; on a shaft that
// crept meanwhile the first VELOCITY command would step by that drift (F324).
// POSITION feeds absolute table values, so only the feed-forward seed applies.
rFeedOn(CLK := bExtWant AND bExtEnabled);
IF rFeedOn.Q THEN
    IF nLoadDomainL = DOM_VELOCITY THEN
        fLoadStartPos := SEL(nLoadMotorL = 1, fLoad2Pos, fLoad1Pos);
        fLoadPosAccum := 0.0;
    END_IF
    fPrevExtPos := SEL(nLoadMotorL = 1, fLoad2Pos, fLoad1Pos);
END_IF

IF bExtWant AND bExtEnabled THEN
    IF nLoadDomainL = DOM_POSITION THEN
        fExtPos := fLoadRaw;                                  // absolute position [deg]
        fExtVel := (fExtPos - fPrevExtPos) / MAX(fDt, 1E-6);  // numeric feed-forward
    ELSE
        fExtPos := fLoadStartPos + fLoadPosAccum;             // VELOCITY: start + integral
        IF eState = ST_RUN THEN fExtVel := fLoadRaw; ELSE fExtVel := 0.0; END_IF
    END_IF
    fPrevExtPos := fExtPos;

    IF   fExtVel > 0.0 THEN nExtDir := 1;
    ELSIF fExtVel < 0.0 THEN nExtDir := -1;
    ELSE                    nExtDir := 0;
    END_IF

    IF nLoadMotorL = 1 THEN
        MC_ExtSetPointGenFeed(Position := fExtPos, Velocity := fExtVel,
                              Acceleration := 0.0, Direction := nExtDir, Axis := AxisLoad1);
    ELSE
        MC_ExtSetPointGenFeed(Position := fExtPos, Velocity := fExtVel,
                              Acceleration := 0.0, Direction := nExtDir, Axis := AxisLoad2);
    END_IF
ELSIF bExtWant THEN
    // engagement pending (standstill wait / sync / enable in flight): scrub
    // the mailbox every cycle so the NC's activation window can only ever
    // see (current actual position, vel 0, Direction 0 = do not apply)
    IF nLoadMotorL = 1 THEN
        MC_ExtSetPointGenFeed(Position := fLoad1Pos, Velocity := 0.0,
                              Acceleration := 0.0, Direction := 0, Axis := AxisLoad1);
    ELSE
        MC_ExtSetPointGenFeed(Position := fLoad2Pos, Velocity := 0.0,
                              Acceleration := 0.0, Direction := 0, Axis := AxisLoad2);
    END_IF
    fPrevExtPos := SEL(nLoadMotorL = 1, fLoad2Pos, fLoad1Pos);
ELSE
    fPrevExtPos := SEL(nLoadMotorL = 1, fLoad2Pos, fLoad1Pos);   // keep the FF seed fresh
END_IF

fbExt1Off(Axis := AxisLoad1, Execute := fExtOff.Q AND (nLoadMotorL = 1));
fbExt2Off(Axis := AxisLoad2, Execute := fExtOff.Q AND (nLoadMotorL = 2));

//----------------------------------------------------------------------
// OUTPUTS / STATUS
//----------------------------------------------------------------------
fMenteeOut           := fMenteeRaw;
fLoadOut             := fLoadRaw;
bRunning             := bWasActive;
stCsv.bRunning       := bRunning;
stCsv.fElapsed       := fElapsed;
stCsv.fMenteeOut     := fMenteeRaw;
stCsv.fLoadOut       := fLoadRaw;
stCsv.bLoadExtActive := bExtWant AND bExtEnabled;

END_FUNCTION_BLOCK

// ---- POUs/FB_HighRateRecorder.TcPOU
// High-rate recorder. Called once per task cycle AFTER the snapshot is assembled.
// While GVL_Recording.bEnable is TRUE it appends one frame to the active chunk of
// GVL_Recording.aChunks (SoA). When a chunk fills it bumps nChunkSeq and advances
// to the next ring slot; the app bulk-reads completed chunks over ADS.
//
// Each frame stores the bus-rate channels (one value) plus the Mentee oversample
// burst (REC_OVERSAMPLE samples). nSampleCount tells the app how many of the
// REC_OVERSAMPLE slots are fresh this frame — the rest are stale (the app keeps
// only the fresh ones and de-dups across frames by sample_idx).
FUNCTION_BLOCK FB_HighRateRecorder
VAR_IN_OUT
    stSnap : ST_SyncSnapshot;   // freshly-assembled snapshot (read only)
END_VAR
VAR
    rEnable : R_TRIG;
    fEnable : F_TRIG;
    nChunk  : UDINT;            // active ring slot (0..REC_RING-1)
    nFill   : UDINT;            // frame index within the active chunk
    nBase   : UDINT;            // Mentee array base = nFill * REC_OVERSAMPLE
    i       : UDINT;
END_VAR

rEnable(CLK := GVL_Recording.bEnable);
fEnable(CLK := GVL_Recording.bEnable);

// Rising edge: start a fresh session (clear ring counters, begin at slot 0).
IF rEnable.Q THEN
    nChunk := 0;
    nFill  := 0;
    GVL_Recording.nChunkSeq := 0;
    GVL_Recording.nReadyIdx := 0;
    GVL_Recording.nDropped  := 0;
    GVL_Recording.nAckSeq   := 0;
    GVL_Recording.aChunks[0].nCount := 0;
    GVL_Recording.bRunning  := TRUE;
END_IF

// Falling edge: flush the partial chunk in progress so the app can capture the
// last (< REC_CHUNK) frames instead of losing them. Publish nFill as nCount and
// bump the sequence exactly like a full chunk; the app honours nCount.
IF fEnable.Q THEN
    GVL_Recording.bRunning := FALSE;
    IF nFill > 0 THEN
        GVL_Recording.aChunks[nChunk].nCount := nFill;
        GVL_Recording.nReadyIdx := TO_BYTE(nChunk);
        GVL_Recording.nChunkSeq := GVL_Recording.nChunkSeq + 1;
        nChunk := (nChunk + 1) MOD GVL_Recording.REC_RING;
        nFill  := 0;
    END_IF
END_IF

IF NOT GVL_Recording.bEnable THEN
    RETURN;
END_IF

// ── append one frame to the active chunk ──
nBase := nFill * GVL_Recording.REC_OVERSAMPLE;

GVL_Recording.aChunks[nChunk].aDcTs[nFill]    := stSnap.nDcTimestamp;
GVL_Recording.aChunks[nChunk].aM1Pos[nFill]   := stSnap.stMotor1Status.fActPosition;
GVL_Recording.aChunks[nChunk].aM1Vel[nFill]   := stSnap.stMotor1Status.fActVelocity;
GVL_Recording.aChunks[nChunk].aM1Trq[nFill]   := stSnap.stMotor1Status.fActTorque;
GVL_Recording.aChunks[nChunk].aM2Pos[nFill]   := stSnap.stMotor2Status.fActPosition;
GVL_Recording.aChunks[nChunk].aM2Vel[nFill]   := stSnap.stMotor2Status.fActVelocity;
GVL_Recording.aChunks[nChunk].aM2Trq[nFill]   := stSnap.stMotor2Status.fActTorque;
GVL_Recording.aChunks[nChunk].aEnc1Cnt[nFill] := stSnap.stEncoder1.nCounterValue;
GVL_Recording.aChunks[nChunk].aEnc1Frq[nFill] := stSnap.stEncoder1.nFrequencyValue;
GVL_Recording.aChunks[nChunk].aEnc2Cnt[nFill] := stSnap.stEncoder2.nCounterValue;
GVL_Recording.aChunks[nChunk].aEnc2Frq[nFill] := stSnap.stEncoder2.nFrequencyValue;
GVL_Recording.aChunks[nChunk].aAin1V[nFill]   := stSnap.stAnalogIn1.fCh1_Voltage;
GVL_Recording.aChunks[nChunk].aAin2V[nFill]   := stSnap.stAnalogIn2.fCh1_Voltage;
GVL_Recording.aChunks[nChunk].aMnSW[nFill]    := stSnap.stMotorV32_OS.nStatusWord;
GVL_Recording.aChunks[nChunk].aMnCnt[nFill]   := stSnap.stMotorV32_OS.nSampleCount;

FOR i := 0 TO GVL_Recording.REC_OVERSAMPLE - 1 DO
    GVL_Recording.aChunks[nChunk].aMnIdx[nBase + i] := stSnap.stMotorV32_OS.aSamples[i].sample_idx;
    GVL_Recording.aChunks[nChunk].aMnW0[nBase + i]  := stSnap.stMotorV32_OS.aSamples[i].w0;
    GVL_Recording.aChunks[nChunk].aMnW1[nBase + i]  := stSnap.stMotorV32_OS.aSamples[i].w1;
    GVL_Recording.aChunks[nChunk].aMnW2[nBase + i]  := stSnap.stMotorV32_OS.aSamples[i].w2;
    // extended lanes 3..9 (ELF-picked debug vars): same slot i, same snapshot,
    // same nBase -> element-aligned with aMnIdx/aMnW0..2 by construction
    GVL_Recording.aChunks[nChunk].aMnW3[nBase + i]  := stSnap.stMotorV32_OS.aSamples[i].w3;
    GVL_Recording.aChunks[nChunk].aMnW4[nBase + i]  := stSnap.stMotorV32_OS.aSamples[i].w4;
    GVL_Recording.aChunks[nChunk].aMnW5[nBase + i]  := stSnap.stMotorV32_OS.aSamples[i].w5;
    GVL_Recording.aChunks[nChunk].aMnW6[nBase + i]  := stSnap.stMotorV32_OS.aSamples[i].w6;
    GVL_Recording.aChunks[nChunk].aMnW7[nBase + i]  := stSnap.stMotorV32_OS.aSamples[i].w7;
    GVL_Recording.aChunks[nChunk].aMnW8[nBase + i]  := stSnap.stMotorV32_OS.aSamples[i].w8;
    GVL_Recording.aChunks[nChunk].aMnW9[nBase + i]  := stSnap.stMotorV32_OS.aSamples[i].w9;
END_FOR

// Futek analog oversamples (EL3702 x5) — raw INT -> V using the same scale as the
// averaged fCh1_Voltage, so the 5 kHz trace is consistent with the 1 kHz average.
FOR i := 1 TO GVL_Recording.REC_FUTEK_OS DO
    GVL_Recording.aChunks[nChunk].aFut1V[nFill * GVL_Recording.REC_FUTEK_OS + (i - 1)] :=
        INT_TO_LREAL(stSnap.stAnalogIn1.nCh1_Sample[i]) / 32767.0 * stSnap.stAnalogIn1.fFullScale;
    GVL_Recording.aChunks[nChunk].aFut2V[nFill * GVL_Recording.REC_FUTEK_OS + (i - 1)] :=
        INT_TO_LREAL(stSnap.stAnalogIn2.nCh1_Sample[i]) / 32767.0 * stSnap.stAnalogIn2.fFullScale;
END_FOR

nFill := nFill + 1;

// ── chunk complete → publish + advance ──
IF nFill >= GVL_Recording.REC_CHUNK THEN
    GVL_Recording.aChunks[nChunk].nCount := GVL_Recording.REC_CHUNK;
    GVL_Recording.nReadyIdx := TO_BYTE(nChunk);
    GVL_Recording.nChunkSeq := GVL_Recording.nChunkSeq + 1;

    // Overflow: the slot we are about to reuse still holds data the app hasn't
    // acked (it is REC_RING-1 chunks behind) — we will overwrite unread data.
    IF (GVL_Recording.nChunkSeq - GVL_Recording.nAckSeq) >= GVL_Recording.REC_RING THEN
        GVL_Recording.nDropped := GVL_Recording.nDropped + GVL_Recording.REC_CHUNK;
    END_IF

    nChunk := (nChunk + 1) MOD GVL_Recording.REC_RING;
    nFill  := 0;
    GVL_Recording.aChunks[nChunk].nCount := 0;   // mark next chunk as "filling"
END_IF

END_FUNCTION_BLOCK

// ---- POUs/FB_UartBridgeHandler.TcPOU
FUNCTION_BLOCK FB_UartBridgeHandler
VAR_IN_OUT
    stCmd               : ST_UartBridgeCmd;
    stStatus            : ST_UartBridgeStatus;
END_VAR

VAR
    //--- RxPDO outputs — AT %Q* — link to device 0x7000 PDOs in XAE ---
    q_control_word      AT %Q* : UDINT; // 0x7000:01 control_word
    q_p_des             AT %Q* : REAL;  // 0x7000:02 p_des
    q_v_des             AT %Q* : REAL;  // 0x7000:03 v_des
    q_kp                AT %Q* : REAL;  // 0x7000:04 kp
    q_kd                AT %Q* : REAL;  // 0x7000:05 kd
    q_torque_ff         AT %Q* : REAL;  // 0x7000:06 torque_ff

    //--- TxPDO inputs — AT %I* — link to device 0x6000 PDOs in XAE ---
    i_status_word       AT %I* : UDINT; // 0x6000:01 status_word
    i_packet_count      AT %I* : UINT;  // 0x6000:02 packet_count
    i_timestamp         AT %I* : UDINT; // 0x6000:03 timestamp
    i_bldc_pos          AT %I* : REAL;  // 0x6000:04 bldc_pos
    i_filtered_p_des    AT %I* : REAL;  // 0x6000:05 filtered_p_des
    i_bldc_vel          AT %I* : REAL;  // 0x6000:06 bldc_vel
    i_v_des             AT %I* : REAL;  // 0x6000:07 v_des
    i_measured_current  AT %I* : REAL;  // 0x6000:08 measured_current
    i_p_i_input         AT %I* : REAL;  // 0x6000:09 p_i_input
    i_impedance_output  AT %I* : REAL;  // 0x6000:0A impedance_output

    //--- Edge detectors for rising edge commands ---
    rtArm           : R_TRIG;
    rtIdle          : R_TRIG;
    rtGateBlock     : R_TRIG;
    rtCalibrate     : R_TRIG;
    rtBode          : R_TRIG;
    rtNoodle        : R_TRIG;
    rtReset         : R_TRIG;
    rtLedOn         : R_TRIG;
    rtLedOff        : R_TRIG;
    rtQueryState    : R_TRIG;

    //--- Internal ---
    nCtrlWord       : UDINT;
END_VAR

//----------------------------------------------------------------------
// EDGE DETECTION — rising edge commands
//----------------------------------------------------------------------
rtArm       (CLK := stCmd.bArm);
rtIdle      (CLK := stCmd.bIdle);
rtGateBlock (CLK := stCmd.bGateBlock);
rtCalibrate (CLK := stCmd.bCalibrate);
rtBode      (CLK := stCmd.bBode);
rtNoodle    (CLK := stCmd.bNoodle);
rtReset     (CLK := stCmd.bReset);
rtLedOn     (CLK := stCmd.bLedOn);
rtLedOff    (CLK := stCmd.bLedOff);
rtQueryState(CLK := stCmd.bQueryState);

//----------------------------------------------------------------------
// BUILD CONTROL WORD
// Rising edge bits — set for one cycle only
// Level bits — held continuously
//----------------------------------------------------------------------
nCtrlWord := 0;

// Rising edge commands — bits 0..9
IF rtArm.Q        THEN nCtrlWord := nCtrlWord OR 16#0001; END_IF
IF rtIdle.Q       THEN nCtrlWord := nCtrlWord OR 16#0002; END_IF
IF rtGateBlock.Q  THEN nCtrlWord := nCtrlWord OR 16#0004; END_IF
IF rtCalibrate.Q  THEN nCtrlWord := nCtrlWord OR 16#0008; END_IF
IF rtBode.Q       THEN nCtrlWord := nCtrlWord OR 16#0010; END_IF
IF rtNoodle.Q     THEN nCtrlWord := nCtrlWord OR 16#0020; END_IF
IF rtReset.Q      THEN nCtrlWord := nCtrlWord OR 16#0040; END_IF
IF rtLedOn.Q      THEN nCtrlWord := nCtrlWord OR 16#0080; END_IF
IF rtLedOff.Q     THEN nCtrlWord := nCtrlWord OR 16#0100; END_IF
IF rtQueryState.Q THEN nCtrlWord := nCtrlWord OR 16#0200; END_IF

// Level: bridge_mode bits 11:10
nCtrlWord := nCtrlWord OR (BYTE_TO_UDINT(stCmd.nBridgeMode AND 16#03) * 16#0400);

// Level: motion_mode bits 14:12
nCtrlWord := nCtrlWord OR (BYTE_TO_UDINT(stCmd.nMotionMode AND 16#07) * 16#1000);

//----------------------------------------------------------------------
// WRITE RxPDO — to device every cycle
//----------------------------------------------------------------------
q_control_word  := nCtrlWord;
q_p_des         := stCmd.p_des;
q_v_des         := stCmd.v_des;
q_kp            := stCmd.kp;
q_kd            := stCmd.kd;
q_torque_ff     := stCmd.torque_ff;

//----------------------------------------------------------------------
// READ TxPDO — from device every cycle
//----------------------------------------------------------------------
stStatus.nStatusWord          := i_status_word;
stStatus.nPacketCount         := i_packet_count;
stStatus.nTimestamp           := i_timestamp;
stStatus.bldc_pos             := i_bldc_pos;
stStatus.filtered_p_des       := i_filtered_p_des;
stStatus.bldc_vel             := i_bldc_vel;
stStatus.v_des                := i_v_des;
stStatus.measured_current     := i_measured_current;
stStatus.p_i_input            := i_p_i_input;
stStatus.impedance_output     := i_impedance_output;

//----------------------------------------------------------------------
// DECODE STATUS WORD
//----------------------------------------------------------------------
stStatus.nFsmState            := UDINT_TO_BYTE(i_status_word AND 16#0000000F);
stStatus.nMainState           := UDINT_TO_BYTE((i_status_word / 16#10)   AND 16#0F);
stStatus.nOpMode              := UDINT_TO_BYTE((i_status_word / 16#100)  AND 16#07);
stStatus.nBridgeModeEcho      := UDINT_TO_BYTE((i_status_word / 16#800)  AND 16#03);
stStatus.nGeneralErrorBits    := UDINT_TO_BYTE((i_status_word / 16#10000) AND 16#FF);
stStatus.nCategorialErrorBits := UDINT_TO_BYTE((i_status_word / 16#1000000) AND 16#FF);
stStatus.bError               := (stStatus.nGeneralErrorBits <> 0)
                               OR (stStatus.nCategorialErrorBits <> 0);

END_FUNCTION_BLOCK

// ---- POUs/CheckBounds.TcPOU
// Implicitly generated code : DO NOT EDIT
FUNCTION CheckBounds : DINT
VAR_INPUT
	index, lower, upper: DINT;
END_VAR
VAR_STAT
	nIndexOverflow : UDINT;
	nIndexUnderflow : UDINT;
END_VAR

// Implicitly generated code: Only an implementation suggestion
{noflow}
IF  index < lower THEN
	nIndexUnderflow := nIndexUnderflow + 1;
	CheckBounds := lower;
ELSIF  index > upper THEN
	nIndexOverflow := nIndexOverflow + 1;
	CheckBounds := upper;
ELSE  
	CheckBounds := index;
END_IF

END_FUNCTION

// ---- POUs/FB_ExtSetpointProbe.TcPOU
// ============================================================================
// FB_ExtSetpointProbe  --  TEMPORARY de-risk probe (delete after verification)
// ----------------------------------------------------------------------------
// Confirms an NC PTP axis accepts EXTERNAL SETPOINT GENERATION (Tc2_MC2):
//   MC_ExtSetPointGenEnable -> MC_ExtSetPointGenFeed (cyclic) -> MC_ExtSetPointGenDisable.
// Setpoints are fed each cycle into Axis.PlcToNc (fExtSetPos/fExtSetVelo/...).
//
// HOW TO RUN (on the bench, motor free / app NOT commanding this axis):
//   1. Instantiate ONE per axis in the active motion program (PRG_Motion):
//        fbProbe1 : FB_ExtSetpointProbe;   // and call fbProbe1(Axis := Axis1);
//      While probing an axis, do NOT also call fbMotor1 for it (two owners
//      of one axis conflict) -- comment that fbMotor call out for the test.
//   2. Set fCycleTime_s to your PLC task period (default 1 ms).
//   3. Online -> write bEnablePower := TRUE, watch bPowered = TRUE.
//   4. Write bRun := TRUE (bFeedSine FALSE). Watch:
//        bExtEnabled = TRUE, bError = FALSE  ==>  EXTERNAL SETPOINT WORKS.
//        bError = TRUE                        ==>  read nErrorID (tells why).
//      (Position is held, so the motor does NOT move in this step.)
//   5. OPTIONAL motion check: write bFeedSine := TRUE -- a slow small sine
//      (fAmplitude / fFrequency) is fed; fActPos should track fSetPos.
//   6. Write bRun := FALSE to hand control back to the NC, then bEnablePower
//      := FALSE. Delete this FB once both axes are confirmed.
// ============================================================================
FUNCTION_BLOCK FB_ExtSetpointProbe
VAR_IN_OUT
    Axis            : AXIS_REF;
END_VAR

VAR_INPUT
    bEnablePower    : BOOL;             // hold TRUE to power the axis (MC_Power)
    bRun            : BOOL;             // TRUE: engage ext-setpoint gen + feed (rising=enable, falling=disable)
    bFeedSine       : BOOL;             // TRUE: feed a slow test sine (MOVES axis); FALSE: hold position
    fAmplitude      : LREAL := 0.5;     // test sine amplitude [axis units]
    fFrequency      : LREAL := 0.2;     // test sine frequency  [Hz]
    fCycleTime_s    : LREAL := 0.001;   // PLC task cycle [s] -- SET to your task period
END_VAR

VAR_OUTPUT
    bPowered        : BOOL;             // MC_Power.Status
    bExtEnabled     : BOOL;             // MC_ExtSetPointGenEnable.Enabled  <-- THE ANSWER
    bError          : BOOL;
    nErrorID        : UDINT;
    fSetPos         : LREAL;            // setpoint position fed (watch vs fActPos)
    fSetVel         : LREAL;            // setpoint velocity fed
    fActPos         : LREAL;            // Axis.NcToPlc.ActPos
END_VAR

VAR
    fbPower         : MC_Power;
    fbExtEnable     : MC_ExtSetPointGenEnable;
    fbExtDisable    : MC_ExtSetPointGenDisable;

    rtRun           : R_TRIG;
    ftRun           : F_TRIG;

    fT              : LREAL;            // elapsed time since enable [s]
    fP0             : LREAL;            // seed position at enable (no jump)
    fW              : LREAL;            // 2*pi*f
    fAcc            : LREAL;            // setpoint acceleration fed
    nDir            : DINT;             // feed direction: 1=+, -1=-, 0=standstill
END_VAR

//----------------------------------------------------------------------
// POWER -- called every cycle
//----------------------------------------------------------------------
fbPower(
    Axis            := Axis,
    Enable          := bEnablePower,
    Enable_Positive := bEnablePower,
    Enable_Negative := bEnablePower,
    Override        := 100.0,
    BufferMode      := MC_Aborting);

rtRun(CLK := bRun);
ftRun(CLK := bRun);

//----------------------------------------------------------------------
// ENABLE external setpoint generation on Run rising edge.
// Seed the profile at the current actual position so there is no jump.
// (Position/PositionType here only arm the optional InTargetPosition
//  monitor; the real setpoints come from MC_ExtSetPointGenFeed below.)
//----------------------------------------------------------------------
IF rtRun.Q THEN
    fP0 := Axis.NcToPlc.ActPos;
    fT  := 0.0;
END_IF

fbExtEnable(
    Axis         := Axis,
    Execute      := rtRun.Q,
    Position     := Axis.NcToPlc.ActPos,
    PositionType := POSITIONTYPE_ABSOLUTE);

//----------------------------------------------------------------------
// FEED the cyclic setpoint while the generator is enabled.
//   bFeedSine = FALSE -> hold fP0 (engage WITHOUT moving the motor).
//   bFeedSine = TRUE  -> slow sine about fP0, with vel/acc feed-forward.
//----------------------------------------------------------------------
IF fbExtEnable.Enabled THEN
    IF bFeedSine THEN
        fT  := fT + fCycleTime_s;
        fW  := 2.0 * 3.14159265358979 * fFrequency;
        fSetPos :=  fP0 + fAmplitude * SIN(fW * fT);
        fSetVel :=  fAmplitude * fW * COS(fW * fT);
        fAcc    := -fAmplitude * fW * fW * SIN(fW * fT);
    ELSE
        fSetPos := fP0;
        fSetVel := 0.0;
        fAcc    := 0.0;
    END_IF

    IF   fSetVel > 0.0 THEN nDir := 1;
    ELSIF fSetVel < 0.0 THEN nDir := -1;
    ELSE                    nDir := 0;
    END_IF

    // Function: copies the values into Axis.PlcToNc (fExtSetPos/Velo/Acc/Dir).
    MC_ExtSetPointGenFeed(
        Position     := fSetPos,
        Velocity     := fSetVel,
        Acceleration := fAcc,
        Direction    := nDir,
        Axis         := Axis);
END_IF

//----------------------------------------------------------------------
// DISABLE on Run falling edge -- hand control back to the NC generator.
//----------------------------------------------------------------------
fbExtDisable(Axis := Axis, Execute := ftRun.Q);

